{region 'Documentation'}
(*!
<summary>Selects literal typed inputs and independent expected results for one comparison row.</summary>
*)
{endregion}
METHOD PRIVATE SelectRow
CASE FRow OF
    BelowZero:
        FActual := LINT#-1;
        FReference := LINT#0;
        FExpectedEqualResult := E_Result.Failed;
        FExpectedNotEqualResult := E_Result.Passed;
        FExpectedLessThanResult := E_Result.Passed;
        FExpectedLessEqualResult := E_Result.Passed;
        FExpectedGreaterThanResult := E_Result.Failed;
        FExpectedGreaterEqualResult := E_Result.Failed;
    EqualZero:
        FActual := LINT#0;
        FReference := LINT#0;
        FExpectedEqualResult := E_Result.Passed;
        FExpectedNotEqualResult := E_Result.Failed;
        FExpectedLessThanResult := E_Result.Failed;
        FExpectedLessEqualResult := E_Result.Passed;
        FExpectedGreaterThanResult := E_Result.Failed;
        FExpectedGreaterEqualResult := E_Result.Passed;
    AboveZero:
        FActual := LINT#1;
        FReference := LINT#0;
        FExpectedEqualResult := E_Result.Failed;
        FExpectedNotEqualResult := E_Result.Passed;
        FExpectedLessThanResult := E_Result.Failed;
        FExpectedLessEqualResult := E_Result.Failed;
        FExpectedGreaterThanResult := E_Result.Passed;
        FExpectedGreaterEqualResult := E_Result.Passed;
    MinimumBelowMaximum:
        FActual := LowestValue;
        FReference := HighestValue;
        FExpectedEqualResult := E_Result.Failed;
        FExpectedNotEqualResult := E_Result.Passed;
        FExpectedLessThanResult := E_Result.Passed;
        FExpectedLessEqualResult := E_Result.Passed;
        FExpectedGreaterThanResult := E_Result.Failed;
        FExpectedGreaterEqualResult := E_Result.Failed;
    MaximumAboveMinimum:
        FActual := HighestValue;
        FReference := LowestValue;
        FExpectedEqualResult := E_Result.Failed;
        FExpectedNotEqualResult := E_Result.Passed;
        FExpectedLessThanResult := E_Result.Failed;
        FExpectedLessEqualResult := E_Result.Failed;
        FExpectedGreaterThanResult := E_Result.Passed;
        FExpectedGreaterEqualResult := E_Result.Passed;
    MinimumEqual:
        FActual := LowestValue;
        FReference := LowestValue;
        FExpectedEqualResult := E_Result.Passed;
        FExpectedNotEqualResult := E_Result.Failed;
        FExpectedLessThanResult := E_Result.Failed;
        FExpectedLessEqualResult := E_Result.Passed;
        FExpectedGreaterThanResult := E_Result.Failed;
        FExpectedGreaterEqualResult := E_Result.Passed;
    MaximumEqual:
        FActual := HighestValue;
        FReference := HighestValue;
        FExpectedEqualResult := E_Result.Passed;
        FExpectedNotEqualResult := E_Result.Failed;
        FExpectedLessThanResult := E_Result.Failed;
        FExpectedLessEqualResult := E_Result.Passed;
        FExpectedGreaterThanResult := E_Result.Failed;
        FExpectedGreaterEqualResult := E_Result.Passed;
ELSE
    Error(Message := 'Unknown comparison test row.');
END_CASE;
END_METHOD

END_FUNCTION_BLOCK

// ---- Framework/Assertions/POU/BasicTypes/LInt/AssertEqual_LInt.TcPOU
{region 'Documentation'}
(*!
<summary>Checks equality with the expected LINT value.</summary>
*)
{endregion}
FUNCTION_BLOCK AssertEqual_LInt EXTENDS AssertionBase
VAR_INPUT
    IN : LINT; //! Actual value checked or observed by this Assertion.
    Expected : LINT; //! Reference value for comparison with IN.
END_VAR

SUPER^();

{region 'Documentation'}
(*!
<summary>Check equality with the expected LINT value.</summary>
*)
{endregion}
METHOD PROTECTED Assert
VAR
    Message : STRING(GVL_Constants.MessageLength);
    ExpectedText : STRING(GVL_Constants.AssertionValueLength);
    ActualText : STRING(GVL_Constants.AssertionValueLength);
END_VAR
IF NOT EvaluationActive THEN
    RETURN;
END_IF;

IF Result = E_Result.Error THEN
    RETURN;
END_IF;

IF Result = E_Result.Failed THEN
    RETURN;
END_IF;

IF IN <> Expected THEN
    ExpectedText := LINT_TO_STRING(Expected);
    ActualText := LINT_TO_STRING(IN);
    Message := CONCAT('Assertion failed: values are not equal. Expected = ',
        ExpectedText);
    Message := CONCAT(Message, ', Actual = ');
    Message := CONCAT(Message, ActualText);
    Message := CONCAT(Message, '.');
    Fail(Message := Message);
    RETURN;
END_IF;

Pass();
END_METHOD

END_FUNCTION_BLOCK

// ---- Framework/Assertions/POU/BasicTypes/LInt/AssertNotEqual_LInt.TcPOU
{region 'Documentation'}
(*!
<summary>Checks inequality with the forbidden LINT value.</summary>
*)
{endregion}
FUNCTION_BLOCK AssertNotEqual_LInt EXTENDS AssertionBase
VAR_INPUT
    IN : LINT; //! Actual value checked or observed by this Assertion.
    Expected : LINT; //! Value that must differ from IN under this Assertion's comparison rules.
END_VAR

SUPER^();

{region 'Documentation'}
(*!
<summary>Check inequality with the forbidden LINT value.</summary>
*)
{endregion}
METHOD PROTECTED Assert
VAR
    Message : STRING(GVL_Constants.MessageLength);
    ExpectedText : STRING(GVL_Constants.AssertionValueLength);
    ActualText : STRING(GVL_Constants.AssertionValueLength);
END_VAR
IF NOT EvaluationActive THEN
    RETURN;
END_IF;

IF Result = E_Result.Error THEN
    RETURN;
END_IF;

IF Result = E_Result.Failed THEN
    RETURN;
END_IF;

IF IN = Expected THEN
    ExpectedText := LINT_TO_STRING(Expected);
    ActualText := LINT_TO_STRING(IN);
    Message := CONCAT('Assertion failed: values are equal but should differ. NotExpected = ',
        ExpectedText);
    Message := CONCAT(Message, ', Actual = ');
    Message := CONCAT(Message, ActualText);
    Message := CONCAT(Message, '.');
    Fail(Message := Message);
    RETURN;
END_IF;

Pass();
END_METHOD

END_FUNCTION_BLOCK

// ---- Framework/Assertions/POU/BasicTypes/LInt/AssertLessThan_LInt.TcPOU
{region 'Documentation'}
(*!
<summary>Check that IN is less than Maximum.</summary>
*)
{endregion}
FUNCTION_BLOCK AssertLessThan_LInt EXTENDS AssertionBase
VAR_INPUT
    IN : LINT; //! Actual value checked or observed by this Assertion.
    Maximum : LINT; //! Exclusive upper bound; the actual value or count must be smaller.
END_VAR

SUPER^();

{region 'Documentation'}
(*!
<summary>Check that IN is less than Maximum.</summary>
*)
{endregion}
METHOD PROTECTED Assert
VAR
    Message : STRING(GVL_Constants.MessageLength);
    MaximumText : STRING(GVL_Constants.AssertionValueLength);
    ActualText : STRING(GVL_Constants.AssertionValueLength);
END_VAR
IF NOT EvaluationActive THEN
    RETURN;
END_IF;

IF Result = E_Result.Error THEN
    RETURN;
END_IF;

IF Result = E_Result.Failed THEN
    RETURN;
END_IF;

IF IN >= Maximum THEN
    MaximumText := LINT_TO_STRING(Maximum);
    ActualText := LINT_TO_STRING(IN);
    Message := CONCAT('Assertion failed: value is not less than maximum. Maximum = ',
        MaximumText);
    Message := CONCAT(Message, ', Actual = ');
    Message := CONCAT(Message, ActualText);
    Message := CONCAT(Message, '.');
    Fail(Message := Message);
    RETURN;
END_IF;

Pass();
END_METHOD

END_FUNCTION_BLOCK

// ---- Framework/Assertions/POU/BasicTypes/LInt/AssertLessEqual_LInt.TcPOU
{region 'Documentation'}
(*!
<summary>Check that IN is at most Maximum.</summary>
*)
{endregion}
FUNCTION_BLOCK AssertLessEqual_LInt EXTENDS AssertionBase
VAR_INPUT
    IN : LINT; //! Actual value checked or observed by this Assertion.
    Maximum : LINT; //! Inclusive upper bound of the comparison; for a range, must not be below Minimum.
END_VAR

SUPER^();

{region 'Documentation'}
(*!
<summary>Check that IN is at most Maximum.</summary>
*)
{endregion}
METHOD PROTECTED Assert
VAR
    Message : STRING(GVL_Constants.MessageLength);
    MaximumText : STRING(GVL_Constants.AssertionValueLength);
    ActualText : STRING(GVL_Constants.AssertionValueLength);
END_VAR
IF NOT EvaluationActive THEN
    RETURN;
END_IF;

IF Result = E_Result.Error THEN
    RETURN;
END_IF;

IF Result = E_Result.Failed THEN
    RETURN;
END_IF;

IF IN > Maximum THEN
    MaximumText := LINT_TO_STRING(Maximum);
    ActualText := LINT_TO_STRING(IN);
    Message := CONCAT('Assertion failed: value is above maximum. Maximum = ',
        MaximumText);
    Message := CONCAT(Message, ', Actual = ');
    Message := CONCAT(Message, ActualText);
    Message := CONCAT(Message, '.');
    Fail(Message := Message);
    RETURN;
END_IF;

Pass();
END_METHOD

END_FUNCTION_BLOCK

// ---- Framework/Assertions/POU/BasicTypes/LInt/AssertGreaterThan_LInt.TcPOU
{region 'Documentation'}
(*!
<summary>Check that IN is greater than Minimum.</summary>
*)
{endregion}
FUNCTION_BLOCK AssertGreaterThan_LInt EXTENDS AssertionBase
VAR_INPUT
    IN : LINT; //! Actual value checked or observed by this Assertion.
    Minimum : LINT; //! Exclusive lower bound; the actual value or count must be greater.
END_VAR

SUPER^();

{region 'Documentation'}
(*!
<summary>Check that IN is greater than Minimum.</summary>
*)
{endregion}
METHOD PROTECTED Assert
VAR
    Message : STRING(GVL_Constants.MessageLength);
    MinimumText : STRING(GVL_Constants.AssertionValueLength);
    ActualText : STRING(GVL_Constants.AssertionValueLength);
END_VAR
IF NOT EvaluationActive THEN
    RETURN;
END_IF;

IF Result = E_Result.Error THEN
    RETURN;
END_IF;

IF Result = E_Result.Failed THEN
    RETURN;
END_IF;

IF IN <= Minimum THEN
    MinimumText := LINT_TO_STRING(Minimum);
    ActualText := LINT_TO_STRING(IN);
    Message := CONCAT('Assertion failed: value is not greater than minimum. Minimum = ',
        MinimumText);
    Message := CONCAT(Message, ', Actual = ');
    Message := CONCAT(Message, ActualText);
    Message := CONCAT(Message, '.');
    Fail(Message := Message);
    RETURN;
END_IF;

Pass();
END_METHOD

END_FUNCTION_BLOCK

// ---- Framework/Assertions/POU/BasicTypes/LInt/AssertGreaterEqual_LInt.TcPOU
{region 'Documentation'}
(*!
<summary>Check that IN is at least Minimum.</summary>
*)
{endregion}
FUNCTION_BLOCK AssertGreaterEqual_LInt EXTENDS AssertionBase
VAR_INPUT
    IN : LINT; //! Actual value checked or observed by this Assertion.
    Minimum : LINT; //! Inclusive lower bound of the comparison; for a range, must not exceed Maximum.
END_VAR

SUPER^();

{region 'Documentation'}
(*!
<summary>Check that IN is at least Minimum.</summary>
*)
{endregion}
METHOD PROTECTED Assert
VAR
    Message : STRING(GVL_Constants.MessageLength);
    MinimumText : STRING(GVL_Constants.AssertionValueLength);
    ActualText : STRING(GVL_Constants.AssertionValueLength);
END_VAR
IF NOT EvaluationActive THEN
    RETURN;
END_IF;

IF Result = E_Result.Error THEN
    RETURN;
END_IF;

IF Result = E_Result.Failed THEN
    RETURN;
END_IF;

IF IN < Minimum THEN
    MinimumText := LINT_TO_STRING(Minimum);
    ActualText := LINT_TO_STRING(IN);
    Message := CONCAT('Assertion failed: value is below minimum. Minimum = ',
        MinimumText);
    Message := CONCAT(Message, ', Actual = ');
    Message := CONCAT(Message, ActualText);
    Message := CONCAT(Message, '.');
    Fail(Message := Message);
    RETURN;
END_IF;

Pass();
END_METHOD

END_FUNCTION_BLOCK

// ---- SelfTests/TestCases/TestSuite_AssertionComparisons/Test_AssertionUnsignedRelations.TcPOU
{region 'Documentation'}
(*!
<summary>Checks six native ULINT comparison relations and full-width boundaries.</summary>
<description>
Each named row has explicit expected results, not a second comparison algorithm.
One disabled subject call consumes Reset before one enabled comparison call.
Outer checking Assertions latch every row before inputs advance; intentional
subject failures remain in a Test-Case-owned Event Buffer, cleared between rows.
Only the checking Assertions contribute to the outer result.
</description>
*)
{endregion}
FUNCTION_BLOCK Test_AssertionUnsignedRelations EXTENDS TestCaseBase
VAR
    FEqualSubject : AssertEqual_ULInt;
    FNotEqualSubject : AssertNotEqual_ULInt;
    FLessThanSubject : AssertLessThan_ULInt;
    FLessEqualSubject : AssertLessEqual_ULInt;
    FGreaterThanSubject : AssertGreaterThan_ULInt;
    FGreaterEqualSubject : AssertGreaterEqual_ULInt;
    FActual : ULINT;
    FReference : ULINT;
    FExpectedEqualResult : E_Result;
    FExpectedNotEqualResult : E_Result;
    FExpectedLessThanResult : E_Result;
    FExpectedLessEqualResult : E_Result;
    FExpectedGreaterThanResult : E_Result;
    FExpectedGreaterEqualResult : E_Result;
    FCapture : EventBuffer;
    FEvents : ARRAY[1..CaptureLength] OF ST_Event;
    FCaptureFifo : ST_FifoStatus;
    FCaptureStatus : ST_EventBufferStatus;
    FRow : UINT;
    FRowPrepared : BOOL;
    FObservationReady : BOOL;
    FChecked : BOOL;
    FSetupValid : BOOL;
END_VAR
VAR
    FEqualResult : AssertTrue;
    FEqualResultMatches : BOOL;
    FNotEqualResult : AssertTrue;
    FNotEqualResultMatches : BOOL;
    FLessThanResult : AssertTrue;
    FLessThanResultMatches : BOOL;
    FLessEqualResult : AssertTrue;
    FLessEqualResultMatches : BOOL;
    FGreaterThanResult : AssertTrue;
    FGreaterThanResultMatches : BOOL;
    FGreaterEqualResult : AssertTrue;
    FGreaterEqualResultMatches : BOOL;
    FCaptureIntegrity : AssertTrue;
    FCaptureIntegrityMatches : BOOL;
END_VAR
VAR CONSTANT
    CaptureLength : UINT := 8;
    ExpectedFindingCount : UDINT := 3;
    BelowSignedBoundary : UINT := 1;
    EqualSignedBoundary : UINT := 2;
    AboveSignedBoundary : UINT := 3;
    ZeroBelowMaximum : UINT := 4;
    MaximumAboveZero : UINT := 5;
    ZeroEqual : UINT := 6;
    MaximumEqual : UINT := 7;
    LastRow : UINT := MaximumEqual;
    SignedBoundary : ULINT := ULINT#9223372036854775808;
    HighestValue : ULINT := ULINT#18446744073709551615;
END_VAR

SUPER^();

{region 'Documentation'}
(*!
<summary>Collects only outer checking Assertions, never intentional subject findings.</summary>
*)
{endregion}
METHOD PROTECTED AggregateResults
VAR_INPUT
    Aggregator : I_ResultAggregator; //! Borrowed result sink owned by the outer Test Case; add this test's checking Assertions without resetting or retaining the sink.
END_VAR
Aggregator.AddProvider(Provider := FEqualResult);
Aggregator.AddProvider(Provider := FNotEqualResult);
Aggregator.AddProvider(Provider := FLessThanResult);
Aggregator.AddProvider(Provider := FLessEqualResult);
Aggregator.AddProvider(Provider := FGreaterThanResult);
Aggregator.AddProvider(Provider := FGreaterEqualResult);
Aggregator.AddProvider(Provider := FCaptureIntegrity);
END_METHOD

{region 'Documentation'}
(*!
<summary>Calls each real comparison once with the selected typed row inputs.</summary>
*)
{endregion}
METHOD PRIVATE CallSubjects
VAR_INPUT
    Enable : BOOL; //! Observation-enable input forwarded to the controlled Assertion subjects for this call.
END_VAR
FEqualSubject(Enable := Enable,
    State := E_State.Running,
    IN := FActual,
    Expected := FReference);
FNotEqualSubject(Enable := Enable,
    State := E_State.Running,
    IN := FActual,
    Expected := FReference);
FLessThanSubject(Enable := Enable,
    State := E_State.Running,
    IN := FActual,
    Maximum := FReference);
FLessEqualSubject(Enable := Enable,
    State := E_State.Running,
    IN := FActual,
    Maximum := FReference);
FGreaterThanSubject(Enable := Enable,
    State := E_State.Running,
    IN := FActual,
    Minimum := FReference);
FGreaterEqualSubject(Enable := Enable,
    State := E_State.Running,
    IN := FActual,
    Minimum := FReference);
END_METHOD

{region 'Documentation'}
(*!
<summary>Preserves base validation and rejects incomplete subject or checking-Assertion setup.</summary>
*)
{endregion}
METHOD PROTECTED CheckInitialization : BOOL //! TRUE when the inherited initialization check and this concrete fixture check both accept the setup.
CheckInitialization := SUPER^.CheckInitialization();
IF NOT CheckInitialization THEN
    RETURN;
END_IF;

CheckInitialization := FSetupValid
    AND FEqualResult.IsInitialized
    AND FNotEqualResult.IsInitialized
    AND FLessThanResult.IsInitialized
    AND FLessEqualResult.IsInitialized
    AND FGreaterThanResult.IsInitialized
    AND FGreaterEqualResult.IsInitialized
    AND FCaptureIntegrity.IsInitialized;
IF NOT CheckInitialization THEN
    EventPublisher.PublishEvent(Event := CreateFrameworkEvent(Name := Name,
        ResourceName := '',
        State := State,
        Severity := E_EventSeverity.Error,
        Message := 'Comparison selftest setup failed.'));
END_IF;
END_METHOD

{region 'Documentation'}
(*!
<summary>Compares observed results with the literal row expectations and checks local event loss/count.</summary>
*)
{endregion}
METHOD PRIVATE CheckResults
FEqualResultMatches := FEqualSubject.Result = FExpectedEqualResult;
FNotEqualResultMatches := FNotEqualSubject.Result = FExpectedNotEqualResult;
FLessThanResultMatches := FLessThanSubject.Result = FExpectedLessThanResult;
FLessEqualResultMatches := FLessEqualSubject.Result = FExpectedLessEqualResult;
FGreaterThanResultMatches := FGreaterThanSubject.Result = FExpectedGreaterThanResult;
FGreaterEqualResultMatches := FGreaterEqualSubject.Result = FExpectedGreaterEqualResult;
FCaptureIntegrityMatches := (FCaptureStatus.SequenceId = ExpectedFindingCount)
    AND (FCaptureStatus.LostEventCount = 0);
END_METHOD

{region 'Documentation'}
(*!
<summary>Initializes the local capture, checking Assertions and publisher-bound real comparisons.</summary>
*)
{endregion}
METHOD PROTECTED Configure
VAR
    Initialized : BOOL;
END_VAR
FPreparationStateCount := 0;
FTestStateCount := 1;
FEqualResult.Initialize(Parent := THIS^,
    AssertionName := 'EqualResult');
FNotEqualResult.Initialize(Parent := THIS^,
    AssertionName := 'NotEqualResult');
FLessThanResult.Initialize(Parent := THIS^,
    AssertionName := 'LessThanResult');
FLessEqualResult.Initialize(Parent := THIS^,
    AssertionName := 'LessEqualResult');
FGreaterThanResult.Initialize(Parent := THIS^,
    AssertionName := 'GreaterThanResult');
FGreaterEqualResult.Initialize(Parent := THIS^,
    AssertionName := 'GreaterEqualResult');
FCaptureIntegrity.Initialize(Parent := THIS^,
    AssertionName := 'CaptureIntegrity');
FSetupValid := FCapture.Initialize(Buffer := FEvents,
    FifoControl := FCaptureFifo,
    Status := FCaptureStatus);
FEqualSubject.BindPublisher(Publisher := FCapture);
Initialized := FEqualSubject.Initialize(Parent := THIS^,
    AssertionName := 'EqualSubject');
FSetupValid := FSetupValid AND Initialized;
FNotEqualSubject.BindPublisher(Publisher := FCapture);
Initialized := FNotEqualSubject.Initialize(Parent := THIS^,
    AssertionName := 'NotEqualSubject');
FSetupValid := FSetupValid AND Initialized;
FLessThanSubject.BindPublisher(Publisher := FCapture);
Initialized := FLessThanSubject.Initialize(Parent := THIS^,
    AssertionName := 'LessThanSubject');
FSetupValid := FSetupValid AND Initialized;
FLessEqualSubject.BindPublisher(Publisher := FCapture);
Initialized := FLessEqualSubject.Initialize(Parent := THIS^,
    AssertionName := 'LessEqualSubject');
FSetupValid := FSetupValid AND Initialized;
FGreaterThanSubject.BindPublisher(Publisher := FCapture);
Initialized := FGreaterThanSubject.Initialize(Parent := THIS^,
    AssertionName := 'GreaterThanSubject');
FSetupValid := FSetupValid AND Initialized;
FGreaterEqualSubject.BindPublisher(Publisher := FCapture);
Initialized := FGreaterEqualSubject.Initialize(Parent := THIS^,
    AssertionName := 'GreaterEqualSubject');
FSetupValid := FSetupValid AND Initialized;
END_METHOD

{region 'Documentation'}
(*!
<summary>Completes abort without asynchronous resources.</summary>
*)
{endregion}
METHOD PROTECTED ProcessAbort
VAR_INPUT
    Enable : BOOL; //! Phase permission supplied by the owning Test Case; FALSE does not authorize progression, while observation may continue.
END_VAR
IF Enable THEN
    CompleteAbort();
END_IF;
END_METHOD

{region 'Documentation'}
(*!
<summary>Latches checked observations before the next script step may proceed.</summary>
*)
{endregion}
METHOD PROTECTED ProcessAssertions
VAR_INPUT
    Enable : BOOL; //! Phase permission supplied by the owning Test Case; FALSE does not authorize progression, while observation may continue.
END_VAR
VAR
    Evaluate : BOOL;
END_VAR
Evaluate := Enable AND FObservationReady;
FEqualResult(Enable := Evaluate,
    State := State,
    IN := FEqualResultMatches);
FNotEqualResult(Enable := Evaluate,
    State := State,
    IN := FNotEqualResultMatches);
FLessThanResult(Enable := Evaluate,
    State := State,
    IN := FLessThanResultMatches);
FLessEqualResult(Enable := Evaluate,
    State := State,
    IN := FLessEqualResultMatches);
FGreaterThanResult(Enable := Evaluate,
    State := State,
    IN := FGreaterThanResultMatches);
FGreaterEqualResult(Enable := Evaluate,
    State := State,
    IN := FGreaterEqualResultMatches);
FCaptureIntegrity(Enable := Evaluate,
    State := State,
    IN := FCaptureIntegrityMatches);
IF Evaluate THEN
    FChecked := TRUE;
END_IF;
END_METHOD

{region 'Documentation'}
(*!
<summary>No Preparation phase is required.</summary>
*)
{endregion}
METHOD PROTECTED ProcessPreparations
VAR_INPUT
    // SA0033: Required hook; this test has no Preparation phase.
    {attribute 'analysis' := '-33'}
    Enable : BOOL; //! Phase permission supplied by the owning Test Case; FALSE does not authorize progression, while observation may continue.
END_VAR
END_METHOD

{region 'Documentation'}
(*!
<summary>Restarts the script and resets the checking Assertions.</summary>
*)
{endregion}
METHOD PROTECTED ProcessReset
FRow := BelowSignedBoundary;
FRowPrepared := FALSE;
FChecked := FALSE;
FObservationReady := FALSE;
FEqualResult.Reset();
FEqualResultMatches := TRUE;
FNotEqualResult.Reset();
FNotEqualResultMatches := TRUE;
FLessThanResult.Reset();
FLessThanResultMatches := TRUE;
FLessEqualResult.Reset();
FLessEqualResultMatches := TRUE;
FGreaterThanResult.Reset();
FGreaterThanResultMatches := TRUE;
FGreaterEqualResult.Reset();
FGreaterEqualResultMatches := TRUE;
FCaptureIntegrity.Reset();
FCaptureIntegrityMatches := TRUE;
CompleteReset();
END_METHOD

{region 'Documentation'}
(*!
<summary>Advances one bounded script step per active PLC cycle.</summary>
*)
{endregion}
METHOD PROTECTED ProcessTests
VAR_INPUT
    Enable : BOOL; //! Phase permission supplied by the owning Test Case; FALSE does not authorize progression, while observation may continue.
END_VAR
IF NOT Enable THEN
    RETURN;
END_IF;

IF FChecked THEN
    FChecked := FALSE;
    FObservationReady := FALSE;
    IF FRow = LastRow THEN
        CompleteTests();
        RETURN;
    END_IF;
    FRow := FRow + 1;
    FRowPrepared := FALSE;
END_IF;

IF NOT FRowPrepared THEN
    SelectRow();
    FCapture.Reset();
    ResetSubjects();
    CallSubjects(Enable := FALSE);
    FRowPrepared := TRUE;
ELSE
    CallSubjects(Enable := TRUE);
    CheckResults();
    FObservationReady := TRUE;
END_IF;
END_METHOD

{region 'Documentation'}
(*!
<summary>Requests a fresh result epoch for every comparison; CallSubjects consumes it.</summary>
*)
{endregion}
METHOD PRIVATE ResetSubjects
FEqualSubject.Reset();
FNotEqualSubject.Reset();
FLessThanSubject.Reset();
FLessEqualSubject.Reset();
FGreaterThanSubject.Reset();
FGreaterEqualSubject.Reset();
END_METHOD

{region 'Documentation'}
(*!
<summary>Selects literal typed inputs and independent expected results for one comparison row.</summary>
*)
{endregion}
METHOD PRIVATE SelectRow
CASE FRow OF
    BelowSignedBoundary:
        FActual := ULINT#9223372036854775807;
        FReference := SignedBoundary;
        FExpectedEqualResult := E_Result.Failed;
        FExpectedNotEqualResult := E_Result.Passed;
        FExpectedLessThanResult := E_Result.Passed;
        FExpectedLessEqualResult := E_Result.Passed;
        FExpectedGreaterThanResult := E_Result.Failed;
        FExpectedGreaterEqualResult := E_Result.Failed;
    EqualSignedBoundary:
        FActual := SignedBoundary;
        FReference := SignedBoundary;
        FExpectedEqualResult := E_Result.Passed;
        FExpectedNotEqualResult := E_Result.Failed;
        FExpectedLessThanResult := E_Result.Failed;
        FExpectedLessEqualResult := E_Result.Passed;
        FExpectedGreaterThanResult := E_Result.Failed;
        FExpectedGreaterEqualResult := E_Result.Passed;
    AboveSignedBoundary:
        FActual := ULINT#9223372036854775809;
        FReference := SignedBoundary;
        FExpectedEqualResult := E_Result.Failed;
        FExpectedNotEqualResult := E_Result.Passed;
        FExpectedLessThanResult := E_Result.Failed;
        FExpectedLessEqualResult := E_Result.Failed;
        FExpectedGreaterThanResult := E_Result.Passed;
        FExpectedGreaterEqualResult := E_Result.Passed;
    ZeroBelowMaximum:
        FActual := ULINT#0;
        FReference := HighestValue;
        FExpectedEqualResult := E_Result.Failed;
        FExpectedNotEqualResult := E_Result.Passed;
        FExpectedLessThanResult := E_Result.Passed;
        FExpectedLessEqualResult := E_Result.Passed;
        FExpectedGreaterThanResult := E_Result.Failed;
        FExpectedGreaterEqualResult := E_Result.Failed;
    MaximumAboveZero:
        FActual := HighestValue;
        FReference := ULINT#0;
        FExpectedEqualResult := E_Result.Failed;
        FExpectedNotEqualResult := E_Result.Passed;
        FExpectedLessThanResult := E_Result.Failed;
        FExpectedLessEqualResult := E_Result.Failed;
        FExpectedGreaterThanResult := E_Result.Passed;
        FExpectedGreaterEqualResult := E_Result.Passed;
    ZeroEqual:
        FActual := ULINT#0;
        FReference := ULINT#0;
        FExpectedEqualResult := E_Result.Passed;
        FExpectedNotEqualResult := E_Result.Failed;
        FExpectedLessThanResult := E_Result.Failed;
        FExpectedLessEqualResult := E_Result.Passed;
        FExpectedGreaterThanResult := E_Result.Failed;
        FExpectedGreaterEqualResult := E_Result.Passed;
    MaximumEqual:
        FActual := HighestValue;
        FReference := HighestValue;
        FExpectedEqualResult := E_Result.Passed;
        FExpectedNotEqualResult := E_Result.Failed;
        FExpectedLessThanResult := E_Result.Failed;
        FExpectedLessEqualResult := E_Result.Passed;
        FExpectedGreaterThanResult := E_Result.Failed;
        FExpectedGreaterEqualResult := E_Result.Passed;
ELSE
    Error(Message := 'Unknown comparison test row.');
END_CASE;
END_METHOD

END_FUNCTION_BLOCK

// ---- SelfTests/TestCases/TestSuite_AssertionComparisons/Test_AssertionBitEquality.TcPOU
{region 'Documentation'}
(*!
<summary>Checks full-value BYTE and LWORD equality without masks or bit-index operations.</summary>
<description>
Each named row has explicit expected results, not a second comparison algorithm.
One disabled subject call consumes Reset before one enabled comparison call.
Outer checking Assertions latch every row before inputs advance; intentional
subject failures remain in a Test-Case-owned Event Buffer, cleared between rows.
Only the checking Assertions contribute to the outer result.
</description>
*)
{endregion}
FUNCTION_BLOCK Test_AssertionBitEquality EXTENDS TestCaseBase
VAR
    FEqualByteSubject : AssertEqual_Byte;
    FNotEqualByteSubject : AssertNotEqual_Byte;
    FEqualLWordSubject : AssertEqual_LWord;
    FNotEqualLWordSubject : AssertNotEqual_LWord;
    FActualByte : BYTE;
    FExpectedByte : BYTE;
    FActualLWord : LWORD;
    FExpectedLWord : LWORD;
    FExpectedEqualByteResult : E_Result;
    FExpectedNotEqualByteResult : E_Result;
    FExpectedEqualLWordResult : E_Result;
    FExpectedNotEqualLWordResult : E_Result;
    FCapture : EventBuffer;
    FEvents : ARRAY[1..CaptureLength] OF ST_Event;
    FCaptureFifo : ST_FifoStatus;
    FCaptureStatus : ST_EventBufferStatus;
    FRow : UINT;
    FRowPrepared : BOOL;
    FObservationReady : BOOL;
    FChecked : BOOL;
    FSetupValid : BOOL;
END_VAR
VAR
    FEqualByteResult : AssertTrue;
    FEqualByteResultMatches : BOOL;
    FNotEqualByteResult : AssertTrue;
    FNotEqualByteResultMatches : BOOL;
    FEqualLWordResult : AssertTrue;
    FEqualLWordResultMatches : BOOL;
    FNotEqualLWordResult : AssertTrue;
    FNotEqualLWordResultMatches : BOOL;
    FCaptureIntegrity : AssertTrue;
    FCaptureIntegrityMatches : BOOL;
END_VAR
VAR CONSTANT
    CaptureLength : UINT := 8;
    ExpectedFindingCount : UDINT := 2;
    ZeroEqual : UINT := 1;
    AllBitsEqual : UINT := 2;
    AllBitsDifferent : UINT := 3;
    HighBitDifferent : UINT := 4;
    PatternDifferent : UINT := 5;
    LastRow : UINT := PatternDifferent;
END_VAR

SUPER^();

{region 'Documentation'}
(*!
<summary>Collects only outer checking Assertions, never intentional subject findings.</summary>
*)
{endregion}
METHOD PROTECTED AggregateResults
VAR_INPUT
    Aggregator : I_ResultAggregator; //! Borrowed result sink owned by the outer Test Case; add this test's checking Assertions without resetting or retaining the sink.
END_VAR
Aggregator.AddProvider(Provider := FEqualByteResult);
Aggregator.AddProvider(Provider := FNotEqualByteResult);
Aggregator.AddProvider(Provider := FEqualLWordResult);
Aggregator.AddProvider(Provider := FNotEqualLWordResult);
Aggregator.AddProvider(Provider := FCaptureIntegrity);
END_METHOD

{region 'Documentation'}
(*!
<summary>Calls each real comparison once with the selected typed row inputs.</summary>
*)
{endregion}
METHOD PRIVATE CallSubjects
VAR_INPUT
    Enable : BOOL; //! Observation-enable input forwarded to the controlled Assertion subjects for this call.
END_VAR
FEqualByteSubject(Enable := Enable,
    State := E_State.Running,
    IN := FActualByte,
    Expected := FExpectedByte);
FNotEqualByteSubject(Enable := Enable,
    State := E_State.Running,
    IN := FActualByte,
    Expected := FExpectedByte);
FEqualLWordSubject(Enable := Enable,
    State := E_State.Running,
    IN := FActualLWord,
    Expected := FExpectedLWord);
FNotEqualLWordSubject(Enable := Enable,
    State := E_State.Running,
    IN := FActualLWord,
    Expected := FExpectedLWord);
END_METHOD

{region 'Documentation'}
(*!
<summary>Preserves base validation and rejects incomplete subject or checking-Assertion setup.</summary>
*)
{endregion}
METHOD PROTECTED CheckInitialization : BOOL //! TRUE when the inherited initialization check and this concrete fixture check both accept the setup.
CheckInitialization := SUPER^.CheckInitialization();
IF NOT CheckInitialization THEN
    RETURN;
END_IF;

CheckInitialization := FSetupValid
    AND FEqualByteResult.IsInitialized
    AND FNotEqualByteResult.IsInitialized
    AND FEqualLWordResult.IsInitialized
    AND FNotEqualLWordResult.IsInitialized
    AND FCaptureIntegrity.IsInitialized;
IF NOT CheckInitialization THEN
    EventPublisher.PublishEvent(Event := CreateFrameworkEvent(Name := Name,
        ResourceName := '',
        State := State,
        Severity := E_EventSeverity.Error,
        Message := 'Comparison selftest setup failed.'));
END_IF;
END_METHOD

{region 'Documentation'}
(*!
<summary>Compares observed results with the literal row expectations and checks local event loss/count.</summary>
*)
{endregion}
METHOD PRIVATE CheckResults
FEqualByteResultMatches := FEqualByteSubject.Result = FExpectedEqualByteResult;
FNotEqualByteResultMatches := FNotEqualByteSubject.Result = FExpectedNotEqualByteResult;
FEqualLWordResultMatches := FEqualLWordSubject.Result = FExpectedEqualLWordResult;
FNotEqualLWordResultMatches := FNotEqualLWordSubject.Result = FExpectedNotEqualLWordResult;
FCaptureIntegrityMatches := (FCaptureStatus.SequenceId = ExpectedFindingCount)
    AND (FCaptureStatus.LostEventCount = 0);
END_METHOD

{region 'Documentation'}
(*!
<summary>Initializes the local capture, checking Assertions and publisher-bound real comparisons.</summary>
*)
{endregion}
METHOD PROTECTED Configure
VAR
    Initialized : BOOL;
END_VAR
FPreparationStateCount := 0;
FTestStateCount := 1;
FEqualByteResult.Initialize(Parent := THIS^,
    AssertionName := 'EqualByteResult');
FNotEqualByteResult.Initialize(Parent := THIS^,
    AssertionName := 'NotEqualByteResult');
FEqualLWordResult.Initialize(Parent := THIS^,
    AssertionName := 'EqualLWordResult');
FNotEqualLWordResult.Initialize(Parent := THIS^,
    AssertionName := 'NotEqualLWordResult');
FCaptureIntegrity.Initialize(Parent := THIS^,
    AssertionName := 'CaptureIntegrity');
FSetupValid := FCapture.Initialize(Buffer := FEvents,
    FifoControl := FCaptureFifo,
    Status := FCaptureStatus);
FEqualByteSubject.BindPublisher(Publisher := FCapture);
Initialized := FEqualByteSubject.Initialize(Parent := THIS^,
    AssertionName := 'EqualByteSubject');
FSetupValid := FSetupValid AND Initialized;
FNotEqualByteSubject.BindPublisher(Publisher := FCapture);
Initialized := FNotEqualByteSubject.Initialize(Parent := THIS^,
    AssertionName := 'NotEqualByteSubject');
FSetupValid := FSetupValid AND Initialized;
FEqualLWordSubject.BindPublisher(Publisher := FCapture);
Initialized := FEqualLWordSubject.Initialize(Parent := THIS^,
    AssertionName := 'EqualLWordSubject');
FSetupValid := FSetupValid AND Initialized;
FNotEqualLWordSubject.BindPublisher(Publisher := FCapture);
Initialized := FNotEqualLWordSubject.Initialize(Parent := THIS^,
    AssertionName := 'NotEqualLWordSubject');
FSetupValid := FSetupValid AND Initialized;
END_METHOD

{region 'Documentation'}
(*!
<summary>Completes abort without asynchronous resources.</summary>
*)
{endregion}
METHOD PROTECTED ProcessAbort
VAR_INPUT
    Enable : BOOL; //! Phase permission supplied by the owning Test Case; FALSE does not authorize progression, while observation may continue.
END_VAR
IF Enable THEN
    CompleteAbort();
END_IF;
END_METHOD

{region 'Documentation'}
(*!
<summary>Latches checked observations before the next script step may proceed.</summary>
*)
{endregion}
METHOD PROTECTED ProcessAssertions
VAR_INPUT
    Enable : BOOL; //! Phase permission supplied by the owning Test Case; FALSE does not authorize progression, while observation may continue.
END_VAR
VAR
    Evaluate : BOOL;
END_VAR
Evaluate := Enable AND FObservationReady;
FEqualByteResult(Enable := Evaluate,
    State := State,
    IN := FEqualByteResultMatches);
FNotEqualByteResult(Enable := Evaluate,
    State := State,
    IN := FNotEqualByteResultMatches);
FEqualLWordResult(Enable := Evaluate,
    State := State,
    IN := FEqualLWordResultMatches);
FNotEqualLWordResult(Enable := Evaluate,
    State := State,
    IN := FNotEqualLWordResultMatches);
FCaptureIntegrity(Enable := Evaluate,
    State := State,
    IN := FCaptureIntegrityMatches);
IF Evaluate THEN
    FChecked := TRUE;
END_IF;
END_METHOD

{region 'Documentation'}
(*!
<summary>No Preparation phase is required.</summary>
*)
{endregion}
METHOD PROTECTED ProcessPreparations
VAR_INPUT
    // SA0033: Required hook; this test has no Preparation phase.
    {attribute 'analysis' := '-33'}
    Enable : BOOL; //! Phase permission supplied by the owning Test Case; FALSE does not authorize progression, while observation may continue.
END_VAR
END_METHOD

{region 'Documentation'}
(*!
<summary>Restarts the script and resets the checking Assertions.</summary>
*)
{endregion}
METHOD PROTECTED ProcessReset
FRow := ZeroEqual;
FRowPrepared := FALSE;
FChecked := FALSE;
FObservationReady := FALSE;
FEqualByteResult.Reset();
FEqualByteResultMatches := TRUE;
FNotEqualByteResult.Reset();
FNotEqualByteResultMatches := TRUE;
FEqualLWordResult.Reset();
FEqualLWordResultMatches := TRUE;
FNotEqualLWordResult.Reset();
FNotEqualLWordResultMatches := TRUE;
FCaptureIntegrity.Reset();
FCaptureIntegrityMatches := TRUE;
CompleteReset();
END_METHOD

{region 'Documentation'}
(*!
<summary>Advances one bounded script step per active PLC cycle.</summary>
*)
{endregion}
METHOD PROTECTED ProcessTests
VAR_INPUT
    Enable : BOOL; //! Phase permission supplied by the owning Test Case; FALSE does not authorize progression, while observation may continue.
END_VAR
IF NOT Enable THEN
    RETURN;
END_IF;

IF FChecked THEN
    FChecked := FALSE;
    FObservationReady := FALSE;
    IF FRow = LastRow THEN
        CompleteTests();
        RETURN;
    END_IF;
    FRow := FRow + 1;
    FRowPrepared := FALSE;
END_IF;

IF NOT FRowPrepared THEN
    SelectRow();
    FCapture.Reset();
    ResetSubjects();
    CallSubjects(Enable := FALSE);
    FRowPrepared := TRUE;
ELSE
    CallSubjects(Enable := TRUE);
    CheckResults();
    FObservationReady := TRUE;
END_IF;
END_METHOD

{region 'Documentation'}
(*!
<summary>Requests a fresh result epoch for every comparison; CallSubjects consumes it.</summary>
*)
{endregion}
METHOD PRIVATE ResetSubjects
FEqualByteSubject.Reset();
FNotEqualByteSubject.Reset();
FEqualLWordSubject.Reset();
FNotEqualLWordSubject.Reset();
END_METHOD

{region 'Documentation'}
(*!
<summary>Selects literal typed inputs and independent expected results for one comparison row.</summary>
*)
{endregion}
METHOD PRIVATE SelectRow
CASE FRow OF
    ZeroEqual:
        FActualByte := BYTE#16#00;
        FExpectedByte := BYTE#16#00;
        FActualLWord := LWORD#16#0000000000000000;
        FExpectedLWord := LWORD#16#0000000000000000;
        FExpectedEqualByteResult := E_Result.Passed;
        FExpectedNotEqualByteResult := E_Result.Failed;
        FExpectedEqualLWordResult := E_Result.Passed;
        FExpectedNotEqualLWordResult := E_Result.Failed;
    AllBitsEqual:
        FActualByte := BYTE#16#FF;
        FExpectedByte := BYTE#16#FF;
        FActualLWord := LWORD#16#FFFFFFFFFFFFFFFF;
        FExpectedLWord := LWORD#16#FFFFFFFFFFFFFFFF;
        FExpectedEqualByteResult := E_Result.Passed;
        FExpectedNotEqualByteResult := E_Result.Failed;
        FExpectedEqualLWordResult := E_Result.Passed;
        FExpectedNotEqualLWordResult := E_Result.Failed;
    AllBitsDifferent:
        FActualByte := BYTE#16#FF;
        FExpectedByte := BYTE#16#00;
        FActualLWord := LWORD#16#FFFFFFFFFFFFFFFF;
        FExpectedLWord := LWORD#16#0000000000000000;
        FExpectedEqualByteResult := E_Result.Failed;
        FExpectedNotEqualByteResult := E_Result.Passed;
        FExpectedEqualLWordResult := E_Result.Failed;
        FExpectedNotEqualLWordResult := E_Result.Passed;
    HighBitDifferent:
        FActualByte := BYTE#16#80;
        FExpectedByte := BYTE#16#00;
        FActualLWord := LWORD#16#8000000000000000;
        FExpectedLWord := LWORD#16#0000000000000000;
        FExpectedEqualByteResult := E_Result.Failed;
        FExpectedNotEqualByteResult := E_Result.Passed;
        FExpectedEqualLWordResult := E_Result.Failed;
        FExpectedNotEqualLWordResult := E_Result.Passed;
    PatternDifferent:
        FActualByte := BYTE#16#A5;
        FExpectedByte := BYTE#16#5A;
        FActualLWord := LWORD#16#A50000000000005A;
        FExpectedLWord := LWORD#16#5A000000000000A5;
        FExpectedEqualByteResult := E_Result.Failed;
        FExpectedNotEqualByteResult := E_Result.Passed;
        FExpectedEqualLWordResult := E_Result.Failed;
        FExpectedNotEqualLWordResult := E_Result.Passed;
ELSE
    Error(Message := 'Unknown comparison test row.');
END_CASE;
END_METHOD

END_FUNCTION_BLOCK

// ---- Framework/Assertions/POU/BasicTypes/Byte/AssertEqual_Byte.TcPOU
{region 'Documentation'}
(*!
<summary>Checks equality with the expected BYTE value.</summary>
*)
{endregion}
FUNCTION_BLOCK AssertEqual_Byte EXTENDS AssertionBase
VAR_INPUT
    IN : BYTE; //! Actual value checked or observed by this Assertion.
    Expected : BYTE; //! Reference value for comparison with IN.
END_VAR

SUPER^();

{region 'Documentation'}
(*!
<summary>Check equality with the expected BYTE value.</summary>
*)
{endregion}
METHOD PROTECTED Assert
VAR
    Message : STRING(GVL_Constants.MessageLength);
    ExpectedText : STRING(GVL_Constants.AssertionValueLength);
    ActualText : STRING(GVL_Constants.AssertionValueLength);
END_VAR
VAR CONSTANT
    HexDigitCount : USINT := 2;
END_VAR
IF NOT EvaluationActive THEN
    RETURN;
END_IF;

IF Result = E_Result.Error THEN
    RETURN;
END_IF;

IF Result = E_Result.Failed THEN
    RETURN;
END_IF;

IF IN <> Expected THEN
    ExpectedText := CreateAssertionTextValue_Hex(Value := BYTE_TO_LWORD(Expected),
        DigitCount := HexDigitCount);
    ActualText := CreateAssertionTextValue_Hex(Value := BYTE_TO_LWORD(IN),
        DigitCount := HexDigitCount);
    Message := CONCAT('Assertion failed: values are not equal. Expected = ',
        ExpectedText);
    Message := CONCAT(Message, ', Actual = ');
    Message := CONCAT(Message, ActualText);
    Message := CONCAT(Message, '.');
    Fail(Message := Message);
    RETURN;
END_IF;

Pass();
END_METHOD

END_FUNCTION_BLOCK

// ---- Framework/Assertions/POU/Utilities/CreateAssertionTextValue_Hex.TcPOU
{region 'Documentation'}
(*!
<summary>Formats a bit-string value as fixed-width uppercase hexadecimal text.</summary>
*)
{endregion}
FUNCTION INTERNAL CreateAssertionTextValue_Hex : STRING(GVL_Constants.AssertionValueLength) //! Bounded diagnostic text; not a value for subsequent numeric comparison.
VAR_INPUT
    Value : LWORD; //! Value to render as diagnostic text; formatting does not change comparison semantics.
    DigitCount : USINT; //! Hexadecimal width, 1..16 digits (2 for BYTE); invalid widths return empty text.
END_VAR
VAR
    RemainingValue : LWORD;
    DigitIndex : INT;
    Nibble : USINT;
    TextValue : STRING(16);
END_VAR
VAR CONSTANT
    HexDigits : STRING(16) := '0123456789ABCDEF';
    MaximumDigits : USINT := 16;
    BitsPerDigit : USINT := 4;
    NibbleMask : LWORD := LWORD#16#F;
END_VAR

IF (DigitCount = 0) OR (DigitCount > MaximumDigits) THEN
    RETURN;
END_IF;

TextValue := '0000000000000000';
// SA0175: DigitCount is 1..16, indices fit STRING(16), masked nibbles are 0..15.
{analysis -175}
TextValue[DigitCount] := 0;
{analysis +175}
RemainingValue := Value;
FOR DigitIndex := USINT_TO_INT(DigitCount) - 1 TO 0 BY -1 DO
    Nibble := LWORD_TO_USINT(RemainingValue AND NibbleMask);
    // SA0175: DigitCount is 1..16, indices fit STRING(16), masked nibbles are 0..15.
    {analysis -175}
    TextValue[DigitIndex] := HexDigits[Nibble];
    {analysis +175}
    RemainingValue := SHR(RemainingValue, BitsPerDigit);
END_FOR;
CreateAssertionTextValue_Hex := CONCAT('16#', TextValue);

END_FUNCTION

// ---- Framework/Assertions/POU/BasicTypes/Byte/AssertNotEqual_Byte.TcPOU
{region 'Documentation'}
(*!
<summary>Checks inequality with the forbidden BYTE value.</summary>
*)
{endregion}
FUNCTION_BLOCK AssertNotEqual_Byte EXTENDS AssertionBase
VAR_INPUT
    IN : BYTE; //! Actual value checked or observed by this Assertion.
    Expected : BYTE; //! Value that must differ from IN under this Assertion's comparison rules.
END_VAR

SUPER^();

{region 'Documentation'}
(*!
<summary>Check inequality with the forbidden BYTE value.</summary>
*)
{endregion}
METHOD PROTECTED Assert
VAR
    Message : STRING(GVL_Constants.MessageLength);
    ExpectedText : STRING(GVL_Constants.AssertionValueLength);
    ActualText : STRING(GVL_Constants.AssertionValueLength);
END_VAR
VAR CONSTANT
    HexDigitCount : USINT := 2;
END_VAR
IF NOT EvaluationActive THEN
    RETURN;
END_IF;

IF Result = E_Result.Error THEN
    RETURN;
END_IF;

IF Result = E_Result.Failed THEN
    RETURN;
END_IF;

IF IN = Expected THEN
    ExpectedText := CreateAssertionTextValue_Hex(Value := BYTE_TO_LWORD(Expected),
        DigitCount := HexDigitCount);
    ActualText := CreateAssertionTextValue_Hex(Value := BYTE_TO_LWORD(IN),
        DigitCount := HexDigitCount);
    Message := CONCAT('Assertion failed: values are equal but should differ. NotExpected = ',
        ExpectedText);
    Message := CONCAT(Message, ', Actual = ');
    Message := CONCAT(Message, ActualText);
    Message := CONCAT(Message, '.');
    Fail(Message := Message);
    RETURN;
END_IF;

Pass();
END_METHOD

END_FUNCTION_BLOCK

// ---- Framework/Assertions/POU/BasicTypes/LWord/AssertEqual_LWord.TcPOU
{region 'Documentation'}
(*!
<summary>Checks equality with the expected LWORD value.</summary>
*)
{endregion}
FUNCTION_BLOCK AssertEqual_LWord EXTENDS AssertionBase
VAR_INPUT
    IN : LWORD; //! Actual value checked or observed by this Assertion.
    Expected : LWORD; //! Reference value for comparison with IN.
END_VAR

SUPER^();

{region 'Documentation'}
(*!
<summary>Check equality with the expected LWORD value.</summary>
*)
{endregion}
METHOD PROTECTED Assert
VAR
    Message : STRING(GVL_Constants.MessageLength);
    ExpectedText : STRING(GVL_Constants.AssertionValueLength);
    ActualText : STRING(GVL_Constants.AssertionValueLength);
END_VAR
VAR CONSTANT
    HexDigitCount : USINT := 16;
END_VAR
IF NOT EvaluationActive THEN
    RETURN;
END_IF;

IF Result = E_Result.Error THEN
    RETURN;
END_IF;

IF Result = E_Result.Failed THEN
    RETURN;
END_IF;

IF IN <> Expected THEN
    ExpectedText := CreateAssertionTextValue_Hex(Value := Expected,
        DigitCount := HexDigitCount);
    ActualText := CreateAssertionTextValue_Hex(Value := IN,
        DigitCount := HexDigitCount);
    Message := CONCAT('Assertion failed: values are not equal. Expected = ',
        ExpectedText);
    Message := CONCAT(Message, ', Actual = ');
    Message := CONCAT(Message, ActualText);
    Message := CONCAT(Message, '.');
    Fail(Message := Message);
    RETURN;
END_IF;

Pass();
END_METHOD

END_FUNCTION_BLOCK

// ---- Framework/Assertions/POU/BasicTypes/LWord/AssertNotEqual_LWord.TcPOU
{region 'Documentation'}
(*!
<summary>Checks inequality with the forbidden LWORD value.</summary>
*)
{endregion}
FUNCTION_BLOCK AssertNotEqual_LWord EXTENDS AssertionBase
VAR_INPUT
    IN : LWORD; //! Actual value checked or observed by this Assertion.
    Expected : LWORD; //! Value that must differ from IN under this Assertion's comparison rules.
END_VAR

SUPER^();

{region 'Documentation'}
(*!
<summary>Check inequality with the forbidden LWORD value.</summary>
*)
{endregion}
METHOD PROTECTED Assert
VAR
    Message : STRING(GVL_Constants.MessageLength);
    ExpectedText : STRING(GVL_Constants.AssertionValueLength);
    ActualText : STRING(GVL_Constants.AssertionValueLength);
END_VAR
VAR CONSTANT
    HexDigitCount : USINT := 16;
END_VAR
IF NOT EvaluationActive THEN
    RETURN;
END_IF;

IF Result = E_Result.Error THEN
    RETURN;
END_IF;

IF Result = E_Result.Failed THEN
    RETURN;
END_IF;

IF IN = Expected THEN
    ExpectedText := CreateAssertionTextValue_Hex(Value := Expected,
        DigitCount := HexDigitCount);
    ActualText := CreateAssertionTextValue_Hex(Value := IN,
        DigitCount := HexDigitCount);
    Message := CONCAT('Assertion failed: values are equal but should differ. NotExpected = ',
        ExpectedText);
    Message := CONCAT(Message, ', Actual = ');
    Message := CONCAT(Message, ActualText);
    Message := CONCAT(Message, '.');
    Fail(Message := Message);
    RETURN;
END_IF;

Pass();
END_METHOD

END_FUNCTION_BLOCK

// ---- SelfTests/TestCases/TestSuite_AssertionComparisons/Test_AssertionBooleanComparisons.TcPOU
{region 'Documentation'}
(*!
<summary>Checks BOOL equality, inequality and direct truth predicates with all truth-table inputs.</summary>
<description>
Each named row has explicit expected results, not a second comparison algorithm.
One disabled subject call consumes Reset before one enabled comparison call.
Outer checking Assertions latch every row before inputs advance; intentional
subject failures remain in a Test-Case-owned Event Buffer, cleared between rows.
Only the checking Assertions contribute to the outer result.
</description>
*)
{endregion}
FUNCTION_BLOCK Test_AssertionBooleanComparisons EXTENDS TestCaseBase
VAR
    FEqualSubject : AssertEqual_Bool;
    FNotEqualSubject : AssertNotEqual_Bool;
    FTrueSubject : AssertTrue;
    FFalseSubject : AssertFalse;
    FActual : BOOL;
    FExpected : BOOL;
    FExpectedEqualResult : E_Result;
    FExpectedNotEqualResult : E_Result;
    FExpectedTrueResult : E_Result;
    FExpectedFalseResult : E_Result;
    FCapture : EventBuffer;
    FEvents : ARRAY[1..CaptureLength] OF ST_Event;
    FCaptureFifo : ST_FifoStatus;
    FCaptureStatus : ST_EventBufferStatus;
    FRow : UINT;
    FRowPrepared : BOOL;
    FObservationReady : BOOL;
    FChecked : BOOL;
    FSetupValid : BOOL;
END_VAR
VAR
    FEqualResult : AssertTrue;
    FEqualResultMatches : BOOL;
    FNotEqualResult : AssertTrue;
    FNotEqualResultMatches : BOOL;
    FTrueResult : AssertTrue;
    FTrueResultMatches : BOOL;
    FFalseResult : AssertTrue;
    FFalseResultMatches : BOOL;
    FCaptureIntegrity : AssertTrue;
    FCaptureIntegrityMatches : BOOL;
END_VAR
VAR CONSTANT
    CaptureLength : UINT := 8;
    ExpectedFindingCount : UDINT := 2;
    BothFalse : UINT := 1;
    FalseVersusTrue : UINT := 2;
    TrueVersusFalse : UINT := 3;
    BothTrue : UINT := 4;
    LastRow : UINT := BothTrue;
END_VAR

SUPER^();

{region 'Documentation'}
(*!
<summary>Collects only outer checking Assertions, never intentional subject findings.</summary>
*)
{endregion}
METHOD PROTECTED AggregateResults
VAR_INPUT
    Aggregator : I_ResultAggregator; //! Borrowed result sink owned by the outer Test Case; add this test's checking Assertions without resetting or retaining the sink.
END_VAR
Aggregator.AddProvider(Provider := FEqualResult);
Aggregator.AddProvider(Provider := FNotEqualResult);
Aggregator.AddProvider(Provider := FTrueResult);
Aggregator.AddProvider(Provider := FFalseResult);
Aggregator.AddProvider(Provider := FCaptureIntegrity);
END_METHOD

{region 'Documentation'}
(*!
<summary>Calls each real comparison once with the selected typed row inputs.</summary>
*)
{endregion}
METHOD PRIVATE CallSubjects
VAR_INPUT
    Enable : BOOL; //! Observation-enable input forwarded to the controlled Assertion subjects for this call.
END_VAR
FEqualSubject(Enable := Enable,
    State := E_State.Running,
    IN := FActual,
    Expected := FExpected);
FNotEqualSubject(Enable := Enable,
    State := E_State.Running,
    IN := FActual,
    Expected := FExpected);
FTrueSubject(Enable := Enable,
    State := E_State.Running,
    IN := FActual);
FFalseSubject(Enable := Enable,
    State := E_State.Running,
    IN := FActual);
END_METHOD

{region 'Documentation'}
(*!
<summary>Preserves base validation and rejects incomplete subject or checking-Assertion setup.</summary>
*)
{endregion}
METHOD PROTECTED CheckInitialization : BOOL //! TRUE when the inherited initialization check and this concrete fixture check both accept the setup.
CheckInitialization := SUPER^.CheckInitialization();
IF NOT CheckInitialization THEN
    RETURN;
END_IF;

CheckInitialization := FSetupValid
    AND FEqualResult.IsInitialized
    AND FNotEqualResult.IsInitialized
    AND FTrueResult.IsInitialized
    AND FFalseResult.IsInitialized
    AND FCaptureIntegrity.IsInitialized;
IF NOT CheckInitialization THEN
    EventPublisher.PublishEvent(Event := CreateFrameworkEvent(Name := Name,
        ResourceName := '',
        State := State,
        Severity := E_EventSeverity.Error,
        Message := 'Comparison selftest setup failed.'));
END_IF;
END_METHOD

{region 'Documentation'}
(*!
<summary>Compares observed results with the literal row expectations and checks local event loss/count.</summary>
*)
{endregion}
METHOD PRIVATE CheckResults
FEqualResultMatches := FEqualSubject.Result = FExpectedEqualResult;
FNotEqualResultMatches := FNotEqualSubject.Result = FExpectedNotEqualResult;
FTrueResultMatches := FTrueSubject.Result = FExpectedTrueResult;
FFalseResultMatches := FFalseSubject.Result = FExpectedFalseResult;
FCaptureIntegrityMatches := (FCaptureStatus.SequenceId = ExpectedFindingCount)
    AND (FCaptureStatus.LostEventCount = 0);
END_METHOD

{region 'Documentation'}
(*!
<summary>Initializes the local capture, checking Assertions and publisher-bound real comparisons.</summary>
*)
{endregion}
METHOD PROTECTED Configure
VAR
    Initialized : BOOL;
END_VAR
FPreparationStateCount := 0;
FTestStateCount := 1;
FEqualResult.Initialize(Parent := THIS^,
    AssertionName := 'EqualResult');
FNotEqualResult.Initialize(Parent := THIS^,
    AssertionName := 'NotEqualResult');
FTrueResult.Initialize(Parent := THIS^,
    AssertionName := 'TrueResult');
FFalseResult.Initialize(Parent := THIS^,
    AssertionName := 'FalseResult');
FCaptureIntegrity.Initialize(Parent := THIS^,
    AssertionName := 'CaptureIntegrity');
FSetupValid := FCapture.Initialize(Buffer := FEvents,
    FifoControl := FCaptureFifo,
    Status := FCaptureStatus);
FEqualSubject.BindPublisher(Publisher := FCapture);
Initialized := FEqualSubject.Initialize(Parent := THIS^,
    AssertionName := 'EqualSubject');
FSetupValid := FSetupValid AND Initialized;
FNotEqualSubject.BindPublisher(Publisher := FCapture);
Initialized := FNotEqualSubject.Initialize(Parent := THIS^,
    AssertionName := 'NotEqualSubject');
FSetupValid := FSetupValid AND Initialized;
FTrueSubject.BindPublisher(Publisher := FCapture);
Initialized := FTrueSubject.Initialize(Parent := THIS^,
    AssertionName := 'TrueSubject');
FSetupValid := FSetupValid AND Initialized;
FFalseSubject.BindPublisher(Publisher := FCapture);
Initialized := FFalseSubject.Initialize(Parent := THIS^,
    AssertionName := 'FalseSubject');
FSetupValid := FSetupValid AND Initialized;
END_METHOD

{region 'Documentation'}
(*!
<summary>Completes abort without asynchronous resources.</summary>
*)
{endregion}
METHOD PROTECTED ProcessAbort
VAR_INPUT
    Enable : BOOL; //! Phase permission supplied by the owning Test Case; FALSE does not authorize progression, while observation may continue.
END_VAR
IF Enable THEN
    CompleteAbort();
END_IF;
END_METHOD

{region 'Documentation'}
(*!
<summary>Latches checked observations before the next script step may proceed.</summary>
*)
{endregion}
METHOD PROTECTED ProcessAssertions
VAR_INPUT
    Enable : BOOL; //! Phase permission supplied by the owning Test Case; FALSE does not authorize progression, while observation may continue.
END_VAR
VAR
    Evaluate : BOOL;
END_VAR
Evaluate := Enable AND FObservationReady;
FEqualResult(Enable := Evaluate,
    State := State,
    IN := FEqualResultMatches);
FNotEqualResult(Enable := Evaluate,
    State := State,
    IN := FNotEqualResultMatches);
FTrueResult(Enable := Evaluate,
    State := State,
    IN := FTrueResultMatches);
FFalseResult(Enable := Evaluate,
    State := State,
    IN := FFalseResultMatches);
FCaptureIntegrity(Enable := Evaluate,
    State := State,
    IN := FCaptureIntegrityMatches);
IF Evaluate THEN
    FChecked := TRUE;
END_IF;
END_METHOD

{region 'Documentation'}
(*!
<summary>No Preparation phase is required.</summary>
*)
{endregion}
METHOD PROTECTED ProcessPreparations
VAR_INPUT
    // SA0033: Required hook; this test has no Preparation phase.
    {attribute 'analysis' := '-33'}
    Enable : BOOL; //! Phase permission supplied by the owning Test Case; FALSE does not authorize progression, while observation may continue.
END_VAR
END_METHOD

{region 'Documentation'}
(*!
<summary>Restarts the script and resets the checking Assertions.</summary>
*)
{endregion}
METHOD PROTECTED ProcessReset
FRow := BothFalse;
FRowPrepared := FALSE;
FChecked := FALSE;
FObservationReady := FALSE;
FEqualResult.Reset();
FEqualResultMatches := TRUE;
FNotEqualResult.Reset();
FNotEqualResultMatches := TRUE;
FTrueResult.Reset();
FTrueResultMatches := TRUE;
FFalseResult.Reset();
FFalseResultMatches := TRUE;
FCaptureIntegrity.Reset();
FCaptureIntegrityMatches := TRUE;
CompleteReset();
END_METHOD

{region 'Documentation'}
(*!
<summary>Advances one bounded script step per active PLC cycle.</summary>
*)
{endregion}
METHOD PROTECTED ProcessTests
VAR_INPUT
    Enable : BOOL; //! Phase permission supplied by the owning Test Case; FALSE does not authorize progression, while observation may continue.
END_VAR
IF NOT Enable THEN
    RETURN;
END_IF;

IF FChecked THEN
    FChecked := FALSE;
    FObservationReady := FALSE;
    IF FRow = LastRow THEN
        CompleteTests();
        RETURN;
    END_IF;
    FRow := FRow + 1;
    FRowPrepared := FALSE;
END_IF;

IF NOT FRowPrepared THEN
    SelectRow();
    FCapture.Reset();
    ResetSubjects();
    CallSubjects(Enable := FALSE);
    FRowPrepared := TRUE;
ELSE
    CallSubjects(Enable := TRUE);
    CheckResults();
    FObservationReady := TRUE;
END_IF;
END_METHOD

{region 'Documentation'}
(*!
<summary>Requests a fresh result epoch for every comparison; CallSubjects consumes it.</summary>
*)
{endregion}
METHOD PRIVATE ResetSubjects
FEqualSubject.Reset();
FNotEqualSubject.Reset();
FTrueSubject.Reset();
FFalseSubject.Reset();
END_METHOD

{region 'Documentation'}
(*!
<summary>Selects literal typed inputs and independent expected results for one comparison row.</summary>
*)
{endregion}
METHOD PRIVATE SelectRow
CASE FRow OF
    BothFalse:
        FActual := FALSE;
        FExpected := FALSE;
        FExpectedEqualResult := E_Result.Passed;
        FExpectedNotEqualResult := E_Result.Failed;
        FExpectedTrueResult := E_Result.Failed;
        FExpectedFalseResult := E_Result.Passed;
    FalseVersusTrue:
        FActual := FALSE;
        FExpected := TRUE;
        FExpectedEqualResult := E_Result.Failed;
        FExpectedNotEqualResult := E_Result.Passed;
        FExpectedTrueResult := E_Result.Failed;
        FExpectedFalseResult := E_Result.Passed;
    TrueVersusFalse:
        FActual := TRUE;
        FExpected := FALSE;
        FExpectedEqualResult := E_Result.Failed;
        FExpectedNotEqualResult := E_Result.Passed;
        FExpectedTrueResult := E_Result.Passed;
        FExpectedFalseResult := E_Result.Failed;
    BothTrue:
        FActual := TRUE;
        FExpected := TRUE;
        FExpectedEqualResult := E_Result.Passed;
        FExpectedNotEqualResult := E_Result.Failed;
        FExpectedTrueResult := E_Result.Passed;
        FExpectedFalseResult := E_Result.Failed;
ELSE
    Error(Message := 'Unknown comparison test row.');
END_CASE;
END_METHOD

END_FUNCTION_BLOCK

// ---- Framework/Assertions/POU/BasicTypes/Bool/AssertNotEqual_Bool.TcPOU
{region 'Documentation'}
(*!
<summary>Checks inequality with the forbidden BOOL value.</summary>
*)
{endregion}
FUNCTION_BLOCK AssertNotEqual_Bool EXTENDS AssertionBase
VAR_INPUT
    IN : BOOL; //! Actual value checked or observed by this Assertion.
    Expected : BOOL; //! Value that must differ from IN under this Assertion's comparison rules.
END_VAR

SUPER^();

{region 'Documentation'}
(*!
<summary>Check inequality with the forbidden BOOL value.</summary>
*)
{endregion}
METHOD PROTECTED Assert
VAR
    Message : STRING(GVL_Constants.MessageLength);
    ExpectedText : STRING(GVL_Constants.AssertionValueLength);
    ActualText : STRING(GVL_Constants.AssertionValueLength);
END_VAR
IF NOT EvaluationActive THEN
    RETURN;
END_IF;

IF Result = E_Result.Error THEN
    RETURN;
END_IF;

IF Result = E_Result.Failed THEN
    RETURN;
END_IF;

IF IN = Expected THEN
    ExpectedText := BOOL_TO_STRING(Expected);
    ActualText := BOOL_TO_STRING(IN);
    Message := CONCAT('Assertion failed: values are equal but should differ. NotExpected = ',
        ExpectedText);
    Message := CONCAT(Message, ', Actual = ');
    Message := CONCAT(Message, ActualText);
    Message := CONCAT(Message, '.');
    Fail(Message := Message);
    RETURN;
END_IF;

Pass();
END_METHOD

END_FUNCTION_BLOCK

// ---- SelfTests/TestCases/TestSuite_AssertionComparisons/Test_AssertionCharacterEquality.TcPOU
{region 'Documentation'}
(*!
<summary>Checks exact BYTE/WORD character-code comparisons for printable, NUL and wide codes.</summary>
<description>
Each named row has explicit expected results, not a second comparison algorithm.
One disabled subject call consumes Reset before one enabled comparison call.
Outer checking Assertions latch every row before inputs advance; intentional
subject failures remain in a Test-Case-owned Event Buffer, cleared between rows.
Only the checking Assertions contribute to the outer result.
</description>
*)
{endregion}
FUNCTION_BLOCK Test_AssertionCharacterEquality EXTENDS TestCaseBase
VAR
    FEqualCharSubject : AssertEqual_Char;
    FNotEqualCharSubject : AssertNotEqual_Char;
    FEqualWCharSubject : AssertEqual_WChar;
    FNotEqualWCharSubject : AssertNotEqual_WChar;
    FActualChar : BYTE;
    FExpectedChar : BYTE;
    FActualWChar : WORD;
    FExpectedWChar : WORD;
    FExpectedEqualCharResult : E_Result;
    FExpectedNotEqualCharResult : E_Result;
    FExpectedEqualWCharResult : E_Result;
    FExpectedNotEqualWCharResult : E_Result;
    FCapture : EventBuffer;
    FEvents : ARRAY[1..CaptureLength] OF ST_Event;
    FCaptureFifo : ST_FifoStatus;
    FCaptureStatus : ST_EventBufferStatus;
    FRow : UINT;
    FRowPrepared : BOOL;
    FObservationReady : BOOL;
    FChecked : BOOL;
    FSetupValid : BOOL;
END_VAR
VAR
    FEqualCharResult : AssertTrue;
    FEqualCharResultMatches : BOOL;
    FNotEqualCharResult : AssertTrue;
    FNotEqualCharResultMatches : BOOL;
    FEqualWCharResult : AssertTrue;
    FEqualWCharResultMatches : BOOL;
    FNotEqualWCharResult : AssertTrue;
    FNotEqualWCharResultMatches : BOOL;
    FCaptureIntegrity : AssertTrue;
    FCaptureIntegrityMatches : BOOL;
END_VAR
VAR CONSTANT
    CaptureLength : UINT := 8;
    ExpectedFindingCount : UDINT := 2;
    PrintableEqual : UINT := 1;
    PrintableDifferent : UINT := 2;
    NullDifferent : UINT := 3;
    NonAsciiDifferent : UINT := 4;
    NullEqual : UINT := 5;
    MaximumEqual : UINT := 6;
    LastRow : UINT := MaximumEqual;
END_VAR

SUPER^();

{region 'Documentation'}
(*!
<summary>Collects only outer checking Assertions, never intentional subject findings.</summary>
*)
{endregion}
METHOD PROTECTED AggregateResults
VAR_INPUT
    Aggregator : I_ResultAggregator; //! Borrowed result sink owned by the outer Test Case; add this test's checking Assertions without resetting or retaining the sink.
END_VAR
Aggregator.AddProvider(Provider := FEqualCharResult);
Aggregator.AddProvider(Provider := FNotEqualCharResult);
Aggregator.AddProvider(Provider := FEqualWCharResult);
Aggregator.AddProvider(Provider := FNotEqualWCharResult);
Aggregator.AddProvider(Provider := FCaptureIntegrity);
END_METHOD

{region 'Documentation'}
(*!
<summary>Calls each real comparison once with the selected typed row inputs.</summary>
*)
{endregion}
METHOD PRIVATE CallSubjects
VAR_INPUT
    Enable : BOOL; //! Observation-enable input forwarded to the controlled Assertion subjects for this call.
END_VAR
FEqualCharSubject(Enable := Enable,
    State := E_State.Running,
    IN := FActualChar,
    Expected := FExpectedChar);
FNotEqualCharSubject(Enable := Enable,
    State := E_State.Running,
    IN := FActualChar,
    Expected := FExpectedChar);
FEqualWCharSubject(Enable := Enable,
    State := E_State.Running,
    IN := FActualWChar,
    Expected := FExpectedWChar);
FNotEqualWCharSubject(Enable := Enable,
    State := E_State.Running,
    IN := FActualWChar,
    Expected := FExpectedWChar);
END_METHOD

{region 'Documentation'}
(*!
<summary>Preserves base validation and rejects incomplete subject or checking-Assertion setup.</summary>
*)
{endregion}
METHOD PROTECTED CheckInitialization : BOOL //! TRUE when the inherited initialization check and this concrete fixture check both accept the setup.
CheckInitialization := SUPER^.CheckInitialization();
IF NOT CheckInitialization THEN
    RETURN;
END_IF;

CheckInitialization := FSetupValid
    AND FEqualCharResult.IsInitialized
    AND FNotEqualCharResult.IsInitialized
    AND FEqualWCharResult.IsInitialized
    AND FNotEqualWCharResult.IsInitialized
    AND FCaptureIntegrity.IsInitialized;
IF NOT CheckInitialization THEN
    EventPublisher.PublishEvent(Event := CreateFrameworkEvent(Name := Name,
        ResourceName := '',
        State := State,
        Severity := E_EventSeverity.Error,
        Message := 'Comparison selftest setup failed.'));
END_IF;
END_METHOD

{region 'Documentation'}
(*!
<summary>Compares observed results with the literal row expectations and checks local event loss/count.</summary>
*)
{endregion}
METHOD PRIVATE CheckResults
FEqualCharResultMatches := FEqualCharSubject.Result = FExpectedEqualCharResult;
FNotEqualCharResultMatches := FNotEqualCharSubject.Result = FExpectedNotEqualCharResult;
FEqualWCharResultMatches := FEqualWCharSubject.Result = FExpectedEqualWCharResult;
FNotEqualWCharResultMatches := FNotEqualWCharSubject.Result = FExpectedNotEqualWCharResult;
FCaptureIntegrityMatches := (FCaptureStatus.SequenceId = ExpectedFindingCount)
    AND (FCaptureStatus.LostEventCount = 0);
END_METHOD

{region 'Documentation'}
(*!
<summary>Initializes the local capture, checking Assertions and publisher-bound real comparisons.</summary>
*)
{endregion}
METHOD PROTECTED Configure
VAR
    Initialized : BOOL;
END_VAR
FPreparationStateCount := 0;
FTestStateCount := 1;
FEqualCharResult.Initialize(Parent := THIS^,
    AssertionName := 'EqualCharResult');
FNotEqualCharResult.Initialize(Parent := THIS^,
    AssertionName := 'NotEqualCharResult');
FEqualWCharResult.Initialize(Parent := THIS^,
    AssertionName := 'EqualWCharResult');
FNotEqualWCharResult.Initialize(Parent := THIS^,
    AssertionName := 'NotEqualWCharResult');
FCaptureIntegrity.Initialize(Parent := THIS^,
    AssertionName := 'CaptureIntegrity');
FSetupValid := FCapture.Initialize(Buffer := FEvents,
    FifoControl := FCaptureFifo,
    Status := FCaptureStatus);
FEqualCharSubject.BindPublisher(Publisher := FCapture);
Initialized := FEqualCharSubject.Initialize(Parent := THIS^,
    AssertionName := 'EqualCharSubject');
FSetupValid := FSetupValid AND Initialized;
FNotEqualCharSubject.BindPublisher(Publisher := FCapture);
Initialized := FNotEqualCharSubject.Initialize(Parent := THIS^,
    AssertionName := 'NotEqualCharSubject');
FSetupValid := FSetupValid AND Initialized;
FEqualWCharSubject.BindPublisher(Publisher := FCapture);
Initialized := FEqualWCharSubject.Initialize(Parent := THIS^,
    AssertionName := 'EqualWCharSubject');
FSetupValid := FSetupValid AND Initialized;
FNotEqualWCharSubject.BindPublisher(Publisher := FCapture);
Initialized := FNotEqualWCharSubject.Initialize(Parent := THIS^,
    AssertionName := 'NotEqualWCharSubject');
FSetupValid := FSetupValid AND Initialized;
END_METHOD

{region 'Documentation'}
(*!
<summary>Completes abort without asynchronous resources.</summary>
*)
{endregion}
METHOD PROTECTED ProcessAbort
VAR_INPUT
    Enable : BOOL; //! Phase permission supplied by the owning Test Case; FALSE does not authorize progression, while observation may continue.
END_VAR
IF Enable THEN
    CompleteAbort();
END_IF;
END_METHOD

{region 'Documentation'}
(*!
<summary>Latches checked observations before the next script step may proceed.</summary>
*)
{endregion}
METHOD PROTECTED ProcessAssertions
VAR_INPUT
    Enable : BOOL; //! Phase permission supplied by the owning Test Case; FALSE does not authorize progression, while observation may continue.
END_VAR
VAR
    Evaluate : BOOL;
END_VAR
Evaluate := Enable AND FObservationReady;
FEqualCharResult(Enable := Evaluate,
    State := State,
    IN := FEqualCharResultMatches);
FNotEqualCharResult(Enable := Evaluate,
    State := State,
    IN := FNotEqualCharResultMatches);
FEqualWCharResult(Enable := Evaluate,
    State := State,
    IN := FEqualWCharResultMatches);
FNotEqualWCharResult(Enable := Evaluate,
    State := State,
    IN := FNotEqualWCharResultMatches);
FCaptureIntegrity(Enable := Evaluate,
    State := State,
    IN := FCaptureIntegrityMatches);
IF Evaluate THEN
    FChecked := TRUE;
END_IF;
END_METHOD

{region 'Documentation'}
(*!
<summary>No Preparation phase is required.</summary>
*)
{endregion}
METHOD PROTECTED ProcessPreparations
VAR_INPUT
    // SA0033: Required hook; this test has no Preparation phase.
    {attribute 'analysis' := '-33'}
    Enable : BOOL; //! Phase permission supplied by the owning Test Case; FALSE does not authorize progression, while observation may continue.
END_VAR
END_METHOD

{region 'Documentation'}
(*!
<summary>Restarts the script and resets the checking Assertions.</summary>
*)
{endregion}
METHOD PROTECTED ProcessReset
FRow := PrintableEqual;
FRowPrepared := FALSE;
FChecked := FALSE;
FObservationReady := FALSE;
FEqualCharResult.Reset();
FEqualCharResultMatches := TRUE;
FNotEqualCharResult.Reset();
FNotEqualCharResultMatches := TRUE;
FEqualWCharResult.Reset();
FEqualWCharResultMatches := TRUE;
FNotEqualWCharResult.Reset();
FNotEqualWCharResultMatches := TRUE;
FCaptureIntegrity.Reset();
FCaptureIntegrityMatches := TRUE;
CompleteReset();
END_METHOD

{region 'Documentation'}
(*!
<summary>Advances one bounded script step per active PLC cycle.</summary>
*)
{endregion}
METHOD PROTECTED ProcessTests
VAR_INPUT
    Enable : BOOL; //! Phase permission supplied by the owning Test Case; FALSE does not authorize progression, while observation may continue.
END_VAR
IF NOT Enable THEN
    RETURN;
END_IF;

IF FChecked THEN
    FChecked := FALSE;
    FObservationReady := FALSE;
    IF FRow = LastRow THEN
        CompleteTests();
        RETURN;
    END_IF;
    FRow := FRow + 1;
    FRowPrepared := FALSE;
END_IF;

IF NOT FRowPrepared THEN
    SelectRow();
    FCapture.Reset();
    ResetSubjects();
    CallSubjects(Enable := FALSE);
    FRowPrepared := TRUE;
ELSE
    CallSubjects(Enable := TRUE);
    CheckResults();
    FObservationReady := TRUE;
END_IF;
END_METHOD

{region 'Documentation'}
(*!
<summary>Requests a fresh result epoch for every comparison; CallSubjects consumes it.</summary>
*)
{endregion}
METHOD PRIVATE ResetSubjects
FEqualCharSubject.Reset();
FNotEqualCharSubject.Reset();
FEqualWCharSubject.Reset();
FNotEqualWCharSubject.Reset();
END_METHOD

{region 'Documentation'}
(*!
<summary>Selects literal typed inputs and independent expected results for one comparison row.</summary>
*)
{endregion}
METHOD PRIVATE SelectRow
CASE FRow OF
    PrintableEqual:
        FActualChar := BYTE#16#41;
        FExpectedChar := BYTE#16#41;
        FActualWChar := WORD#16#0041;
        FExpectedWChar := WORD#16#0041;
        FExpectedEqualCharResult := E_Result.Passed;
        FExpectedNotEqualCharResult := E_Result.Failed;
        FExpectedEqualWCharResult := E_Result.Passed;
        FExpectedNotEqualWCharResult := E_Result.Failed;
    PrintableDifferent:
        FActualChar := BYTE#16#41;
        FExpectedChar := BYTE#16#42;
        FActualWChar := WORD#16#0041;
        FExpectedWChar := WORD#16#0042;
        FExpectedEqualCharResult := E_Result.Failed;
        FExpectedNotEqualCharResult := E_Result.Passed;
        FExpectedEqualWCharResult := E_Result.Failed;
        FExpectedNotEqualWCharResult := E_Result.Passed;
    NullDifferent:
        FActualChar := BYTE#16#00;
        FExpectedChar := BYTE#16#41;
        FActualWChar := WORD#16#0000;
        FExpectedWChar := WORD#16#0041;
        FExpectedEqualCharResult := E_Result.Failed;
        FExpectedNotEqualCharResult := E_Result.Passed;
        FExpectedEqualWCharResult := E_Result.Failed;
        FExpectedNotEqualWCharResult := E_Result.Passed;
    NonAsciiDifferent:
        FActualChar := BYTE#16#FF;
        FExpectedChar := BYTE#16#41;
        FActualWChar := WORD#16#0100;
        FExpectedWChar := WORD#16#0000;
        FExpectedEqualCharResult := E_Result.Failed;
        FExpectedNotEqualCharResult := E_Result.Passed;
        FExpectedEqualWCharResult := E_Result.Failed;
        FExpectedNotEqualWCharResult := E_Result.Passed;
    NullEqual:
        FActualChar := BYTE#16#00;
        FExpectedChar := BYTE#16#00;
        FActualWChar := WORD#16#0000;
        FExpectedWChar := WORD#16#0000;
        FExpectedEqualCharResult := E_Result.Passed;
        FExpectedNotEqualCharResult := E_Result.Failed;
        FExpectedEqualWCharResult := E_Result.Passed;
        FExpectedNotEqualWCharResult := E_Result.Failed;
    MaximumEqual:
        FActualChar := BYTE#16#FF;
        FExpectedChar := BYTE#16#FF;
        FActualWChar := WORD#16#FFFF;
        FExpectedWChar := WORD#16#FFFF;
        FExpectedEqualCharResult := E_Result.Passed;
        FExpectedNotEqualCharResult := E_Result.Failed;
        FExpectedEqualWCharResult := E_Result.Passed;
        FExpectedNotEqualWCharResult := E_Result.Failed;
ELSE
    Error(Message := 'Unknown comparison test row.');
END_CASE;
END_METHOD

END_FUNCTION_BLOCK

// ---- Framework/Assertions/POU/BasicTypes/Char/AssertEqual_Char.TcPOU
{region 'Documentation'}
(*!
<summary>Checks exact equality of character codes.</summary>
<description>

Character codes use BYTE; diagnostics show printable ASCII and hexadecimal codes.

Compares the numeric character code without case folding or encoding validation.
Printable ASCII diagnostics include the character and hexadecimal code; other codes use a
hexadecimal representation.

</description>
*)
{endregion}
FUNCTION_BLOCK AssertEqual_Char EXTENDS AssertionBase
VAR_INPUT
    IN : BYTE; //! Actual character code.
    Expected : BYTE; //! Expected character code.
END_VAR

SUPER^();

{region 'Documentation'}
(*!
<summary>Compares character codes and reports character-formatted diagnostics.</summary>
*)
{endregion}
METHOD PROTECTED Assert
VAR
    Message : STRING(GVL_Constants.MessageLength);
    ExpectedText : STRING;
    ActualText : STRING;
END_VAR
IF NOT EvaluationActive THEN
    RETURN;
END_IF;

IF Result = E_Result.Error THEN
    RETURN;
END_IF;

IF Result = E_Result.Failed THEN
    RETURN;
END_IF;

IF IN <> Expected THEN
    ExpectedText := CreateAssertionTextValue_Char(Value := Expected);
    ActualText := CreateAssertionTextValue_Char(Value := IN);
    Message := CONCAT('Assertion failed: values are not equal. Expected = ',
        ExpectedText);
    Message := CONCAT(Message, ', Actual = ');
    Message := CONCAT(Message, ActualText);
    Message := CONCAT(Message, '.');
    Fail(Message := Message);
    RETURN;
END_IF;

Pass();
END_METHOD

END_FUNCTION_BLOCK

// ---- Framework/Assertions/POU/Utilities/CreateAssertionTextValue_Char.TcPOU
{region 'Documentation'}
(*!
<summary>Formats printable ASCII as a quoted character and hexadecimal code; other values as code only. Output is ASCII and at most 11 characters.</summary>
*)
{endregion}
FUNCTION INTERNAL CreateAssertionTextValue_Char : STRING(11) //! Bounded diagnostic text; not a value for subsequent numeric comparison.
VAR_INPUT
    Value : BYTE; //! Character code to render; no character validation is performed.
END_VAR
VAR
    HexText : STRING(5);
    Text : STRING(11);
END_VAR
VAR CONSTANT
    FirstPrintableAscii : BYTE := 16#20;
    LastPrintableAscii : BYTE := 16#7E;
    HexDigitCount : USINT := 2;
END_VAR

HexText := CreateAssertionTextValue_Hex(Value := BYTE_TO_LWORD(Value),
    DigitCount := HexDigitCount);

IF (Value < FirstPrintableAscii) OR (Value > LastPrintableAscii) THEN
    CreateAssertionTextValue_Char := HexText;
    RETURN;
END_IF;

Text := '$' $' (';
// SA0175: Printable-ASCII guard; index 1 fits the quoted template.
{analysis -175}
Text[1] := Value;
{analysis +175}
Text := CONCAT(Text, HexText);
CreateAssertionTextValue_Char := CONCAT(Text, ')');

END_FUNCTION

// ---- Framework/Assertions/POU/BasicTypes/Char/AssertNotEqual_Char.TcPOU
{region 'Documentation'}
(*!
<summary>Checks exact inequality of character codes.</summary>
<description>

Character codes use BYTE; diagnostics show printable ASCII and hexadecimal codes.

Compares the numeric character code without case folding or encoding validation.
Printable ASCII diagnostics include the character and hexadecimal code; other codes use a
hexadecimal representation.

</description>
*)
{endregion}
FUNCTION_BLOCK AssertNotEqual_Char EXTENDS AssertionBase
VAR_INPUT
    IN : BYTE; //! Actual character code.
    Expected : BYTE; //! Forbidden character code.
END_VAR

SUPER^();

{region 'Documentation'}
(*!
<summary>Compares character codes and reports character-formatted diagnostics.</summary>
*)
{endregion}
METHOD PROTECTED Assert
VAR
    Message : STRING(GVL_Constants.MessageLength);
    ExpectedText : STRING;
    ActualText : STRING;
END_VAR
IF NOT EvaluationActive THEN
    RETURN;
END_IF;

IF Result = E_Result.Error THEN
    RETURN;
END_IF;

IF Result = E_Result.Failed THEN
    RETURN;
END_IF;

IF IN = Expected THEN
    ExpectedText := CreateAssertionTextValue_Char(Value := Expected);
    ActualText := CreateAssertionTextValue_Char(Value := IN);
    Message := CONCAT('Assertion failed: values are equal. NotExpected = ',
        ExpectedText);
    Message := CONCAT(Message, ', Actual = ');
    Message := CONCAT(Message, ActualText);
    Message := CONCAT(Message, '.');
    Fail(Message := Message);
    RETURN;
END_IF;

Pass();
END_METHOD

END_FUNCTION_BLOCK

// ---- SelfTests/TestCases/TestSuite_AssertionComparisons/Test_AssertionSignedRanges.TcPOU
{region 'Documentation'}
(*!
<summary>Checks inclusive LINT ranges, reversed bounds and Failed-to-Error escalation.</summary>
<description>
Named rows separate independent comparisons by a disabled reset call.
Only explicitly marked escalation rows retain the preceding subject result.
Outer Assertions latch every observation before advancing to the next row.
Intentional findings remain in the local capture; no production algorithm is copied.
</description>
*)
{endregion}
FUNCTION_BLOCK Test_AssertionSignedRanges EXTENDS TestCaseBase
VAR
    FInRangeSubject : AssertInRange_LInt;
    FNotInRangeSubject : AssertNotInRange_LInt;
    FActual : LINT;
    FLower : LINT;
    FUpper : LINT;
    FExpectedInRangeResult : E_Result;
    FExpectedNotInRangeResult : E_Result;
    FExpectedFindings : UDINT;
    FCapture : EventBuffer;
    FEvents : ARRAY[1..CaptureLength] OF ST_Event;
    FCaptureFifo : ST_FifoStatus;
    FCaptureStatus : ST_EventBufferStatus;
    FRow : UINT;
    FRowPrepared : BOOL;
    FPreserveResults : BOOL;
    FObservationReady : BOOL;
    FChecked : BOOL;
    FSetupValid : BOOL;
END_VAR
VAR
    FInRangeResult : AssertTrue;
    FInRangeResultMatches : BOOL;
    FNotInRangeResult : AssertTrue;
    FNotInRangeResultMatches : BOOL;
    FCaptureIntegrity : AssertTrue;
    FCaptureIntegrityMatches : BOOL;
END_VAR
VAR CONSTANT
    CaptureLength : UINT := 8;
    LowerEndpoint : UINT := 1;
    Interior : UINT := 2;
    UpperEndpoint : UINT := 3;
    BelowRange : UINT := 4;
    AboveRange : UINT := 5;
    EqualBounds : UINT := 6;
    ReversedBounds : UINT := 7;
    MinimumEndpoint : UINT := 8;
    MaximumEndpoint : UINT := 9;
    FailureBeforeInvalid : UINT := 10;
    InvalidAfterFailure : UINT := 11;
    LastRow : UINT := InvalidAfterFailure;
    LowestValue : LINT := LINT#-9223372036854775808;
    HighestValue : LINT := LINT#9223372036854775807;
END_VAR

SUPER^();

{region 'Documentation'}
(*!
<summary>Collects only outer checking Assertions, never intentional subject findings.</summary>
*)
{endregion}
METHOD PROTECTED AggregateResults
VAR_INPUT
    Aggregator : I_ResultAggregator; //! Borrowed result sink owned by the outer Test Case; add this test's checking Assertions without resetting or retaining the sink.
END_VAR
Aggregator.AddProvider(Provider := FInRangeResult);
Aggregator.AddProvider(Provider := FNotInRangeResult);
Aggregator.AddProvider(Provider := FCaptureIntegrity);
END_METHOD

{region 'Documentation'}
(*!
<summary>Calls each inherited production Assertion once using the selected row.</summary>
*)
{endregion}
METHOD PRIVATE CallSubjects
VAR_INPUT
    Enable : BOOL; //! Observation-enable input forwarded to the controlled Assertion subjects for this call.
END_VAR
FInRangeSubject(Enable := Enable,
    State := E_State.Running,
    IN := FActual,
    Minimum := FLower,
    Maximum := FUpper);
FNotInRangeSubject(Enable := Enable,
    State := E_State.Running,
    IN := FActual,
    Minimum := FLower,
    Maximum := FUpper);
END_METHOD

{region 'Documentation'}
(*!
<summary>Extends base validation with subject and checking-Assertion setup.</summary>
*)
{endregion}
METHOD PROTECTED CheckInitialization : BOOL //! TRUE when the inherited initialization check and this concrete fixture check both accept the setup.
CheckInitialization := SUPER^.CheckInitialization();
IF NOT CheckInitialization THEN
    RETURN;
END_IF;

CheckInitialization := FSetupValid
    AND FInRangeResult.IsInitialized
    AND FNotInRangeResult.IsInitialized
    AND FCaptureIntegrity.IsInitialized;
IF NOT CheckInitialization THEN
    EventPublisher.PublishEvent(Event := CreateFrameworkEvent(Name := Name,
        ResourceName := '',
        State := State,
        Severity := E_EventSeverity.Error,
        Message := 'Comparison selftest setup failed.'));
END_IF;
END_METHOD

{region 'Documentation'}
(*!
<summary>Checks results and isolated findings against explicit expectations.</summary>
*)
{endregion}
METHOD PRIVATE CheckResults
FInRangeResultMatches := FInRangeSubject.Result = FExpectedInRangeResult;
FNotInRangeResultMatches := FNotInRangeSubject.Result = FExpectedNotInRangeResult;
FCaptureIntegrityMatches := (FCaptureStatus.SequenceId = FExpectedFindings)
    AND (FCaptureStatus.LostEventCount = 0);
END_METHOD

{region 'Documentation'}
(*!
<summary>Configures checking Assertions; subject actions remain in the test script.</summary>
*)
{endregion}
METHOD PROTECTED Configure
VAR
    Initialized : BOOL;
END_VAR
FPreparationStateCount := 0;
FTestStateCount := 1;
FInRangeResult.Initialize(Parent := THIS^,
    AssertionName := 'InRangeResult');
FNotInRangeResult.Initialize(Parent := THIS^,
    AssertionName := 'NotInRangeResult');
FCaptureIntegrity.Initialize(Parent := THIS^,
    AssertionName := 'CaptureIntegrity');
FSetupValid := FCapture.Initialize(Buffer := FEvents,
    FifoControl := FCaptureFifo,
    Status := FCaptureStatus);
FInRangeSubject.BindPublisher(Publisher := FCapture);
Initialized := FInRangeSubject.Initialize(Parent := THIS^,
    AssertionName := 'InRangeSubject');
FSetupValid := FSetupValid AND Initialized;
FNotInRangeSubject.BindPublisher(Publisher := FCapture);
Initialized := FNotInRangeSubject.Initialize(Parent := THIS^,
    AssertionName := 'NotInRangeSubject');
FSetupValid := FSetupValid AND Initialized;
END_METHOD

{region 'Documentation'}
(*!
<summary>Completes abort without asynchronous resources.</summary>
*)
{endregion}
METHOD PROTECTED ProcessAbort
VAR_INPUT
    Enable : BOOL; //! Phase permission supplied by the owning Test Case; FALSE does not authorize progression, while observation may continue.
END_VAR
IF Enable THEN
    CompleteAbort();
END_IF;
END_METHOD

{region 'Documentation'}
(*!
<summary>Latches checked observations before the next script step may proceed.</summary>
*)
{endregion}
METHOD PROTECTED ProcessAssertions
VAR_INPUT
    Enable : BOOL; //! Phase permission supplied by the owning Test Case; FALSE does not authorize progression, while observation may continue.
END_VAR
VAR
    Evaluate : BOOL;
END_VAR
Evaluate := Enable AND FObservationReady;
FInRangeResult(Enable := Evaluate,
    State := State,
    IN := FInRangeResultMatches);
FNotInRangeResult(Enable := Evaluate,
    State := State,
    IN := FNotInRangeResultMatches);
FCaptureIntegrity(Enable := Evaluate,
    State := State,
    IN := FCaptureIntegrityMatches);
IF Evaluate THEN
    FChecked := TRUE;
END_IF;
END_METHOD

{region 'Documentation'}
(*!
<summary>No Preparation phase is required.</summary>
*)
{endregion}
METHOD PROTECTED ProcessPreparations
VAR_INPUT
    // SA0033: Required hook; this test has no Preparation phase.
    {attribute 'analysis' := '-33'}
    Enable : BOOL; //! Phase permission supplied by the owning Test Case; FALSE does not authorize progression, while observation may continue.
END_VAR
END_METHOD

{region 'Documentation'}
(*!
<summary>Restarts the script and resets the checking Assertions.</summary>
*)
{endregion}
METHOD PROTECTED ProcessReset
FRow := LowerEndpoint;
FRowPrepared := FALSE;
FChecked := FALSE;
FObservationReady := FALSE;
FInRangeResult.Reset();
FInRangeResultMatches := TRUE;
FNotInRangeResult.Reset();
FNotInRangeResultMatches := TRUE;
FCaptureIntegrity.Reset();
FCaptureIntegrityMatches := TRUE;
CompleteReset();
END_METHOD

{region 'Documentation'}
(*!
<summary>Advances one bounded script step per active PLC cycle.</summary>
*)
{endregion}
METHOD PROTECTED ProcessTests
VAR_INPUT
    Enable : BOOL; //! Phase permission supplied by the owning Test Case; FALSE does not authorize progression, while observation may continue.
END_VAR
IF NOT Enable THEN
    RETURN;
END_IF;

IF FChecked THEN
    FChecked := FALSE;
    FObservationReady := FALSE;
    IF FRow = LastRow THEN
        CompleteTests();
        RETURN;
    END_IF;
    FRow := FRow + 1;
    FRowPrepared := FALSE;
END_IF;

IF NOT FRowPrepared THEN
    SelectRow();
    FCapture.Reset();
    IF NOT FPreserveResults THEN
        ResetSubjects();
    END_IF;
    CallSubjects(Enable := FALSE);
    FRowPrepared := TRUE;
ELSE
    CallSubjects(Enable := TRUE);
    CheckResults();
    FObservationReady := TRUE;
END_IF;
END_METHOD

{region 'Documentation'}
(*!
<summary>Requests fresh subject results before the next disabled call.</summary>
*)
{endregion}
METHOD PRIVATE ResetSubjects
FInRangeSubject.Reset();
FNotInRangeSubject.Reset();
END_METHOD

{region 'Documentation'}
(*!
<summary>Selects literal expectations; only named escalation rows retain preceding subject results.</summary>
*)
{endregion}
METHOD PRIVATE SelectRow
FPreserveResults := FALSE;
CASE FRow OF
    LowerEndpoint:
        FActual := LINT#-1;
        FLower := LINT#-1;
        FUpper := LINT#1;
        FExpectedInRangeResult := E_Result.Passed;
        FExpectedNotInRangeResult := E_Result.Failed;
        FExpectedFindings := 1;
    Interior:
        FActual := LINT#0;
        FLower := LINT#-1;
        FUpper := LINT#1;
        FExpectedInRangeResult := E_Result.Passed;
        FExpectedNotInRangeResult := E_Result.Failed;
        FExpectedFindings := 1;
    UpperEndpoint:
        FActual := LINT#1;
        FLower := LINT#-1;
        FUpper := LINT#1;
        FExpectedInRangeResult := E_Result.Passed;
        FExpectedNotInRangeResult := E_Result.Failed;
        FExpectedFindings := 1;
    BelowRange:
        FActual := LINT#-2;
        FLower := LINT#-1;
        FUpper := LINT#1;
        FExpectedInRangeResult := E_Result.Failed;
        FExpectedNotInRangeResult := E_Result.Passed;
        FExpectedFindings := 1;
    AboveRange:
        FActual := LINT#2;
        FLower := LINT#-1;
        FUpper := LINT#1;
        FExpectedInRangeResult := E_Result.Failed;
        FExpectedNotInRangeResult := E_Result.Passed;
        FExpectedFindings := 1;
    EqualBounds:
        FActual := LINT#0;
        FLower := LINT#0;
        FUpper := LINT#0;
        FExpectedInRangeResult := E_Result.Passed;
        FExpectedNotInRangeResult := E_Result.Failed;
        FExpectedFindings := 1;
    ReversedBounds:
        FActual := LINT#0;
        FLower := LINT#1;
        FUpper := LINT#-1;
        FExpectedInRangeResult := E_Result.Error;
        FExpectedNotInRangeResult := E_Result.Error;
        FExpectedFindings := 2;
    MinimumEndpoint:
        FActual := LowestValue;
        FLower := LowestValue;
        FUpper := HighestValue;
        FExpectedInRangeResult := E_Result.Passed;
        FExpectedNotInRangeResult := E_Result.Failed;
        FExpectedFindings := 1;
    MaximumEndpoint:
        FActual := HighestValue;
        FLower := LowestValue;
        FUpper := HighestValue;
        FExpectedInRangeResult := E_Result.Passed;
        FExpectedNotInRangeResult := E_Result.Failed;
        FExpectedFindings := 1;
    FailureBeforeInvalid:
        FActual := LINT#2;
        FLower := LINT#-1;
        FUpper := LINT#1;
        FExpectedInRangeResult := E_Result.Failed;
        FExpectedNotInRangeResult := E_Result.Passed;
        FExpectedFindings := 1;
    InvalidAfterFailure:
        FActual := LINT#0;
        FLower := LINT#1;
        FUpper := LINT#-1;
        FExpectedInRangeResult := E_Result.Error;
        FExpectedNotInRangeResult := E_Result.Error;
        FExpectedFindings := 2;
        FPreserveResults := TRUE;
ELSE
    Error(Message := 'Unknown comparison test row.');
END_CASE;
END_METHOD

END_FUNCTION_BLOCK

// ---- Framework/Assertions/POU/BasicTypes/LInt/AssertInRange_LInt.TcPOU
{region 'Documentation'}
(*!
<summary>Checks whether the LINT value is inside the inclusive range.</summary>
<description>

Minimum &gt; Maximum reports Error during active evaluation; equal bounds are
valid.

</description>
*)
{endregion}
FUNCTION_BLOCK AssertInRange_LInt EXTENDS AssertionBase
VAR_INPUT
    IN : LINT; //! Actual value checked or observed by this Assertion.
    Minimum : LINT; //! Inclusive lower bound of the comparison; for a range, must not exceed Maximum.
    Maximum : LINT; //! Inclusive upper bound of the comparison; for a range, must not be below Minimum.
END_VAR

SUPER^();

{region 'Documentation'}
(*!
<summary>Check whether the LINT value is inside the inclusive range.</summary>
*)
{endregion}
METHOD PROTECTED Assert
VAR
    Message : STRING(GVL_Constants.MessageLength);
    MinimumText : STRING(GVL_Constants.AssertionValueLength);
    MaximumText : STRING(GVL_Constants.AssertionValueLength);
    ActualText : STRING(GVL_Constants.AssertionValueLength);
END_VAR
IF NOT EvaluationActive THEN
    RETURN;
END_IF;

IF Result = E_Result.Error THEN
    RETURN;
END_IF;

IF Minimum > Maximum THEN
    MinimumText := LINT_TO_STRING(Minimum);
    MaximumText := LINT_TO_STRING(Maximum);
    Message := CONCAT('Assertion error: minimum exceeds maximum. Minimum = ',
        MinimumText);
    Message := CONCAT(Message, ', Maximum = ');
    Message := CONCAT(Message, MaximumText);
    Message := CONCAT(Message, '.');
    Error(Message := Message);
    RETURN;
END_IF;

IF Result = E_Result.Failed THEN
    RETURN;
END_IF;

IF (IN < Minimum) OR (IN > Maximum) THEN
    MinimumText := LINT_TO_STRING(Minimum);
    MaximumText := LINT_TO_STRING(Maximum);
    ActualText := LINT_TO_STRING(IN);
    Message := CONCAT('Assertion failed: value is outside allowed range. Minimum = ',
        MinimumText);
    Message := CONCAT(Message, ', Maximum = ');
    Message := CONCAT(Message, MaximumText);
    Message := CONCAT(Message, ', Actual = ');
    Message := CONCAT(Message, ActualText);
    Message := CONCAT(Message, '.');
    Fail(Message := Message);
    RETURN;
END_IF;

Pass();
END_METHOD

END_FUNCTION_BLOCK

// ---- Framework/Assertions/POU/BasicTypes/LInt/AssertNotInRange_LInt.TcPOU
{region 'Documentation'}
(*!
<summary>Checks whether the LINT value is outside the inclusive range.</summary>
<description>

Minimum &gt; Maximum reports Error during active evaluation; equal bounds are
valid.

</description>
*)
{endregion}
FUNCTION_BLOCK AssertNotInRange_LInt EXTENDS AssertionBase
VAR_INPUT
    IN : LINT; //! Actual value checked or observed by this Assertion.
    Minimum : LINT; //! Inclusive lower bound of the comparison; for a range, must not exceed Maximum.
    Maximum : LINT; //! Inclusive upper bound of the comparison; for a range, must not be below Minimum.
END_VAR

SUPER^();

{region 'Documentation'}
(*!
<summary>Check whether the LINT value is outside the inclusive range.</summary>
*)
{endregion}
METHOD PROTECTED Assert
VAR
    Message : STRING(GVL_Constants.MessageLength);
    MinimumText : STRING(GVL_Constants.AssertionValueLength);
    MaximumText : STRING(GVL_Constants.AssertionValueLength);
    ActualText : STRING(GVL_Constants.AssertionValueLength);
END_VAR
IF NOT EvaluationActive THEN
    RETURN;
END_IF;

IF Result = E_Result.Error THEN
    RETURN;
END_IF;

IF Minimum > Maximum THEN
    MinimumText := LINT_TO_STRING(Minimum);
    MaximumText := LINT_TO_STRING(Maximum);
    Message := CONCAT('Assertion error: minimum exceeds maximum. Minimum = ',
        MinimumText);
    Message := CONCAT(Message, ', Maximum = ');
    Message := CONCAT(Message, MaximumText);
    Message := CONCAT(Message, '.');
    Error(Message := Message);
    RETURN;
END_IF;

IF Result = E_Result.Failed THEN
    RETURN;
END_IF;

IF (IN >= Minimum) AND (IN <= Maximum) THEN
    MinimumText := LINT_TO_STRING(Minimum);
    MaximumText := LINT_TO_STRING(Maximum);
    ActualText := LINT_TO_STRING(IN);
    Message := CONCAT('Assertion failed: value is inside forbidden range. Minimum = ',
        MinimumText);
    Message := CONCAT(Message, ', Maximum = ');
    Message := CONCAT(Message, MaximumText);
    Message := CONCAT(Message, ', Actual = ');
    Message := CONCAT(Message, ActualText);
    Message := CONCAT(Message, '.');
    Fail(Message := Message);
    RETURN;
END_IF;

Pass();
END_METHOD

END_FUNCTION_BLOCK

// ---- SelfTests/TestCases/TestSuite_AssertionComparisons/Test_AssertionUnsignedRanges.TcPOU
{region 'Documentation'}
(*!
<summary>Checks inclusive ULINT ranges, reversed bounds and Failed-to-Error escalation.</summary>
<description>
Named rows separate independent comparisons by a disabled reset call.
Only explicitly marked escalation rows retain the preceding subject result.
Outer Assertions latch every observation before advancing to the next row.
Intentional findings remain in the local capture; no production algorithm is copied.
</description>
*)
{endregion}
FUNCTION_BLOCK Test_AssertionUnsignedRanges EXTENDS TestCaseBase
VAR
    FInRangeSubject : AssertInRange_ULInt;
    FNotInRangeSubject : AssertNotInRange_ULInt;
    FActual : ULINT;
    FLower : ULINT;
    FUpper : ULINT;
    FExpectedInRangeResult : E_Result;
    FExpectedNotInRangeResult : E_Result;
    FExpectedFindings : UDINT;
    FCapture : EventBuffer;
    FEvents : ARRAY[1..CaptureLength] OF ST_Event;
    FCaptureFifo : ST_FifoStatus;
    FCaptureStatus : ST_EventBufferStatus;
    FRow : UINT;
    FRowPrepared : BOOL;
    FPreserveResults : BOOL;
    FObservationReady : BOOL;
    FChecked : BOOL;
    FSetupValid : BOOL;
END_VAR
VAR
    FInRangeResult : AssertTrue;
    FInRangeResultMatches : BOOL;
    FNotInRangeResult : AssertTrue;
    FNotInRangeResultMatches : BOOL;
    FCaptureIntegrity : AssertTrue;
    FCaptureIntegrityMatches : BOOL;
END_VAR
VAR CONSTANT
    CaptureLength : UINT := 8;
    LowerEndpoint : UINT := 1;
    Interior : UINT := 2;
    UpperEndpoint : UINT := 3;
    BelowRange : UINT := 4;
    AboveRange : UINT := 5;
    EqualBounds : UINT := 6;
    ReversedBounds : UINT := 7;
    MinimumEndpoint : UINT := 8;
    MaximumEndpoint : UINT := 9;
    FailureBeforeInvalid : UINT := 10;
    InvalidAfterFailure : UINT := 11;
    LastRow : UINT := InvalidAfterFailure;
    LowestValue : ULINT := ULINT#0;
    HighestValue : ULINT := ULINT#18446744073709551615;
END_VAR

SUPER^();

{region 'Documentation'}
(*!
<summary>Collects only outer checking Assertions, never intentional subject findings.</summary>
*)
{endregion}
METHOD PROTECTED AggregateResults
VAR_INPUT
    Aggregator : I_ResultAggregator; //! Borrowed result sink owned by the outer Test Case; add this test's checking Assertions without resetting or retaining the sink.
END_VAR
Aggregator.AddProvider(Provider := FInRangeResult);
Aggregator.AddProvider(Provider := FNotInRangeResult);
Aggregator.AddProvider(Provider := FCaptureIntegrity);
END_METHOD

{region 'Documentation'}
(*!
<summary>Calls each inherited production Assertion once using the selected row.</summary>
*)
{endregion}
METHOD PRIVATE CallSubjects
VAR_INPUT
    Enable : BOOL; //! Observation-enable input forwarded to the controlled Assertion subjects for this call.
END_VAR
FInRangeSubject(Enable := Enable,
    State := E_State.Running,
    IN := FActual,
    Minimum := FLower,
    Maximum := FUpper);
FNotInRangeSubject(Enable := Enable,
    State := E_State.Running,
    IN := FActual,
    Minimum := FLower,
    Maximum := FUpper);
END_METHOD

{region 'Documentation'}
(*!
<summary>Extends base validation with subject and checking-Assertion setup.</summary>
*)
{endregion}
METHOD PROTECTED CheckInitialization : BOOL //! TRUE when the inherited initialization check and this concrete fixture check both accept the setup.
CheckInitialization := SUPER^.CheckInitialization();
IF NOT CheckInitialization THEN
    RETURN;
END_IF;

CheckInitialization := FSetupValid
    AND FInRangeResult.IsInitialized
    AND FNotInRangeResult.IsInitialized
    AND FCaptureIntegrity.IsInitialized;
IF NOT CheckInitialization THEN
    EventPublisher.PublishEvent(Event := CreateFrameworkEvent(Name := Name,
        ResourceName := '',
        State := State,
        Severity := E_EventSeverity.Error,
        Message := 'Comparison selftest setup failed.'));
END_IF;
END_METHOD

{region 'Documentation'}
(*!
<summary>Checks results and isolated findings against explicit expectations.</summary>
*)
{endregion}
METHOD PRIVATE CheckResults
FInRangeResultMatches := FInRangeSubject.Result = FExpectedInRangeResult;
FNotInRangeResultMatches := FNotInRangeSubject.Result = FExpectedNotInRangeResult;
FCaptureIntegrityMatches := (FCaptureStatus.SequenceId = FExpectedFindings)
    AND (FCaptureStatus.LostEventCount = 0);
END_METHOD

{region 'Documentation'}
(*!
<summary>Configures checking Assertions; subject actions remain in the test script.</summary>
*)
{endregion}
METHOD PROTECTED Configure
VAR
    Initialized : BOOL;
END_VAR
FPreparationStateCount := 0;
FTestStateCount := 1;
FInRangeResult.Initialize(Parent := THIS^,
    AssertionName := 'InRangeResult');
FNotInRangeResult.Initialize(Parent := THIS^,
    AssertionName := 'NotInRangeResult');
FCaptureIntegrity.Initialize(Parent := THIS^,
    AssertionName := 'CaptureIntegrity');
FSetupValid := FCapture.Initialize(Buffer := FEvents,
    FifoControl := FCaptureFifo,
    Status := FCaptureStatus);
FInRangeSubject.BindPublisher(Publisher := FCapture);
Initialized := FInRangeSubject.Initialize(Parent := THIS^,
    AssertionName := 'InRangeSubject');
FSetupValid := FSetupValid AND Initialized;
FNotInRangeSubject.BindPublisher(Publisher := FCapture);
Initialized := FNotInRangeSubject.Initialize(Parent := THIS^,
    AssertionName := 'NotInRangeSubject');
FSetupValid := FSetupValid AND Initialized;
END_METHOD

{region 'Documentation'}
(*!
<summary>Completes abort without asynchronous resources.</summary>
*)
{endregion}
METHOD PROTECTED ProcessAbort
VAR_INPUT
    Enable : BOOL; //! Phase permission supplied by the owning Test Case; FALSE does not authorize progression, while observation may continue.
END_VAR
IF Enable THEN
    CompleteAbort();
END_IF;
END_METHOD

{region 'Documentation'}
(*!
<summary>Latches checked observations before the next script step may proceed.</summary>
*)
{endregion}
METHOD PROTECTED ProcessAssertions
VAR_INPUT
    Enable : BOOL; //! Phase permission supplied by the owning Test Case; FALSE does not authorize progression, while observation may continue.
END_VAR
VAR
    Evaluate : BOOL;
END_VAR
Evaluate := Enable AND FObservationReady;
FInRangeResult(Enable := Evaluate,
    State := State,
    IN := FInRangeResultMatches);
FNotInRangeResult(Enable := Evaluate,
    State := State,
    IN := FNotInRangeResultMatches);
FCaptureIntegrity(Enable := Evaluate,
    State := State,
    IN := FCaptureIntegrityMatches);
IF Evaluate THEN
    FChecked := TRUE;
END_IF;
END_METHOD

{region 'Documentation'}
(*!
<summary>No Preparation phase is required.</summary>
*)
{endregion}
METHOD PROTECTED ProcessPreparations
VAR_INPUT
    // SA0033: Required hook; this test has no Preparation phase.
    {attribute 'analysis' := '-33'}
    Enable : BOOL; //! Phase permission supplied by the owning Test Case; FALSE does not authorize progression, while observation may continue.
END_VAR
END_METHOD

{region 'Documentation'}
(*!
<summary>Restarts the script and resets the checking Assertions.</summary>
*)
{endregion}
METHOD PROTECTED ProcessReset
FRow := LowerEndpoint;
FRowPrepared := FALSE;
FChecked := FALSE;
FObservationReady := FALSE;
FInRangeResult.Reset();
FInRangeResultMatches := TRUE;
FNotInRangeResult.Reset();
FNotInRangeResultMatches := TRUE;
FCaptureIntegrity.Reset();
FCaptureIntegrityMatches := TRUE;
CompleteReset();
END_METHOD

{region 'Documentation'}
(*!
<summary>Advances one bounded script step per active PLC cycle.</summary>
*)
{endregion}
METHOD PROTECTED ProcessTests
VAR_INPUT
    Enable : BOOL; //! Phase permission supplied by the owning Test Case; FALSE does not authorize progression, while observation may continue.
END_VAR
IF NOT Enable THEN
    RETURN;
END_IF;

IF FChecked THEN
    FChecked := FALSE;
    FObservationReady := FALSE;
    IF FRow = LastRow THEN
        CompleteTests();
        RETURN;
    END_IF;
    FRow := FRow + 1;
    FRowPrepared := FALSE;
END_IF;

